(* IEC 61131-3 sources: daoli-st-library/DL_Motion (part 17) *)

(* ---- FB_DL_ServoVelLoopBand.st ---- *)
(* ===========================================================================
   组件名   : FB_DL_ServoVelLoopBand
   分类     : DL_Motion / 速度环带宽估算
   一句话   : 由速度指令阶跃响应的 10%→90% 上升时间估算闭环带宽并判定是否达标
   复杂度   : 2        版本 : v1.0.0        日期 : 2026-11-24
   开源溯源 : 无（clean-room 自研，未借鉴任何开源实现）
   输入契约 : xEnable 功能使能；xArm 测量许可（FALSE 复位）；fVelRef 速度指令 [rpm]
              fVelFbk 速度反馈 [rpm]；fDtSec 采样周期 [s]；fStepThr 阶跃识别阈值 [rpm]
              fRiseLowFrac/fRiseHighFrac 上升时间取点分数；fTimeoutSec 测量超时 [s]
              fBandFactor 上升时间-带宽系数（一阶近似 0.35）；fBandTargetHz 达标带宽 [Hz]
   输出契约 : fRiseTimeSec 上升时间 [s]；fBandwidthHz 估算带宽 [Hz]；xDone 测量完成
              xBandOk 带宽达标（容差比较）；xValid 输入有效
              iErrorCode 0=正常 1=输入非有限 2=测量超时 3=上升时间过小 9=非法状态
   修改记录 : v1.0.0 2026-11-24 初版
   =========================================================================== *)

TYPE E_DL_RiseMeasState :
(
    eIdle := 0,       // 空闲待命 | idle
    eWaitStep := 1,   // 等待阶跃发生 | wait for step
    eRising := 2,     // 上升沿测量中 | rising measurement
    eDone := 3,       // 测量完成 | measurement done
    eFail := 4        // 测量失败 | measurement failed
);
END_TYPE

FUNCTION_BLOCK FB_DL_ServoVelLoopBand
VAR_INPUT
    xEnable : BOOL;                       // 功能使能 | function enable
    xArm : BOOL;                          // 测量许可 FALSE=复位 | measurement arm
    fVelRef : REAL;                       // 速度指令 [rpm] | velocity reference [rpm]
    fVelFbk : REAL;                       // 速度反馈 [rpm] | velocity feedback [rpm]
    fDtSec : REAL := 0.004;               // 采样周期 [s] | sample period [s]
    fStepThr : REAL := 50.0;              // 阶跃识别阈值 [rpm] | step detect threshold [rpm]
    fRiseLowFrac : REAL := 0.1;           // 上升时间起点分数 | rise time low fraction
    fRiseHighFrac : REAL := 0.9;          // 上升时间终点分数 | rise time high fraction
    fTimeoutSec : REAL := 5.0;            // 测量超时 [s] | measurement timeout [s]
    fBandFactor : REAL := 0.35;           // 上升时间-带宽系数 | rise time band factor
    fBandTargetHz : REAL := 100.0;        // 达标带宽 [Hz] | target bandwidth [Hz]
END_VAR
VAR_OUTPUT
    fRiseTimeSec : REAL;                  // 上升时间 [s] | rise time [s]
    fBandwidthHz : REAL;                  // 估算带宽 [Hz] | estimated bandwidth [Hz]
    xDone : BOOL;                         // 测量完成 | measurement done
    xBandOk : BOOL;                       // 带宽达标 | bandwidth acceptable
    xValid : BOOL;                        // 输入有效标志 | inputs valid flag
    iErrorCode : INT;                     // 故障码 0=无故障 | error code
    eStateOut : E_DL_RiseMeasState;       // 当前状态观测 | current state observation
END_VAR
VAR
    _eState : E_DL_RiseMeasState := eIdle;  // 内部状态机状态 | internal state
    _fRefPrev : REAL;                     // 上一拍速度指令 [rpm] | previous reference [rpm]
    _fStart : REAL;                       // 阶跃起点值 [rpm] | step start value [rpm]
    _fAmp : REAL;                         // 阶跃幅值 [rpm] | step amplitude [rpm]
    _fElapsed : REAL;                     // 阶跃后累计时间 [s] | elapsed since step [s]
    _fProg : REAL;                        // 归一化响应进度 | normalized response progress
    _fT10 : REAL;                         // 10% 时刻 [s] | time at low fraction [s]
    _fT90 : REAL;                         // 90% 时刻 [s] | time at high fraction [s]
    _fDt : REAL;                          // 钳位后采样周期 [s] | clamped dt [s]
    _xGot10 : BOOL;                       // 已捕获低分数时刻 | low fraction captured
    _xGot90 : BOOL;                       // 已捕获高分数时刻 | high fraction captured
    _xBad : BOOL;                         // 输入非有限标志 | not-finite flag
    _xBadPar : BOOL;                      // 参数非法标志 | invalid parameter flag
END_VAR

// ---- 非有限检测 ----
_xBad := (fVelRef <> fVelRef) OR ((fVelRef - fVelRef) <> (fVelRef - fVelRef))
      OR (fVelFbk <> fVelFbk) OR ((fVelFbk - fVelFbk) <> (fVelFbk - fVelFbk))
      OR (fDtSec <> fDtSec) OR ((fDtSec - fDtSec) <> (fDtSec - fDtSec))
      OR (fBandFactor <> fBandFactor) OR ((fBandFactor - fBandFactor) <> (fBandFactor - fBandFactor));

// ---- 参数合法性：所有做分母/做取点的量必须为正且分数有序 ----
_xBadPar := (fDtSec <= 0.0) OR (fStepThr <= 0.0) OR (fTimeoutSec <= 0.0)
         OR (fBandFactor <= 0.0) OR (fBandTargetHz <= 0.0)
         OR (fRiseLowFrac <= 0.0) OR (fRiseHighFrac <= fRiseLowFrac);

xValid := NOT (_xBad OR _xBadPar);
iErrorCode := 0;
IF _xBad THEN
    iErrorCode := 1;
ELSIF _xBadPar THEN
    iErrorCode := 2;
END_IF

// ---- 周期钳位 ----
_fDt := fDtSec;
IF _fDt < 0.000001 THEN
    _fDt := 0.000001;
ELSIF _fDt > 0.2 THEN
    _fDt := 0.2;
END_IF

CASE _eState OF
    eIdle:
        xDone := FALSE;
        IF NOT xEnable THEN
            iErrorCode := 0;
        ELSIF xArm AND xValid THEN
            fRiseTimeSec := 0.0;
            fBandwidthHz := 0.0;
            xBandOk := FALSE;
            _fElapsed := 0.0;
            _eState := eWaitStep;
        END_IF

    eWaitStep:
        IF NOT xArm OR NOT xEnable THEN
            _eState := eIdle;
        ELSIF ABS(fVelRef - _fRefPrev) > fStepThr THEN
            _fStart := _fRefPrev;                    // 阶跃起点
            _fAmp := fVelRef - _fRefPrev;            // 阶跃幅值
            IF ABS(_fAmp) > 0.000000001 THEN          // 防零除：幅值必须显著
                _fElapsed := 0.0;
                _fT10 := 0.0;
                _fT90 := 0.0;
                _xGot10 := FALSE;
                _xGot90 := FALSE;
                _eState := eRising;
            ELSE
                iErrorCode := 3;                     // 幅值过小视为无效阶跃
                _eState := eFail;
            END_IF
        END_IF

    eRising:
        IF NOT xArm OR NOT xEnable THEN
            _eState := eIdle;
        ELSE
            _fElapsed := _fElapsed + _fDt;
            _fProg := 0.0;
            IF ABS(_fAmp) > 0.000000001 THEN
                _fProg := (fVelFbk - _fStart) / _fAmp;   // 归一化进度，分母已守卫
            END_IF
            IF NOT _xGot10 AND (_fProg >= fRiseLowFrac) THEN
                _fT10 := _fElapsed;
                _xGot10 := TRUE;
            END_IF
            IF _xGot10 AND NOT _xGot90 AND (_fProg >= fRiseHighFrac) THEN
                _fT90 := _fElapsed;
                _xGot90 := TRUE;
            END_IF
            IF _xGot90 THEN
                fRiseTimeSec := _fT90 - _fT10;
                IF fRiseTimeSec > 0.000001 THEN
                    fBandwidthHz := fBandFactor / fRiseTimeSec;   // 分母已守卫
                    xDone := TRUE;
                    _eState := eDone;
                ELSE
                    iErrorCode := 3;                 // 上升时间过小，估算不可信
                    _eState := eFail;
                END_IF
            ELSIF _fElapsed > fTimeoutSec THEN
                iErrorCode := 2;                     // 响应未达 90%，测量超时
                _eState := eFail;
            END_IF
        END_IF

    eDone:
        IF NOT xArm OR NOT xEnable THEN
            xDone := FALSE;
            _eState := eIdle;                        // 结果保持至下一次重新测量
        END_IF

    eFail:
        xDone := FALSE;
        IF NOT xArm OR NOT xEnable THEN
            iErrorCode := 0;
            _eState := eIdle;
        END_IF

ELSE
    iErrorCode := 9;                                 // 非法状态兜底
    xDone := FALSE;
    _eState := eIdle;
END_CASE;

// ---- 达标判定：仅在测量完成后用容差比较带宽 ----
IF _eState = eDone THEN
    xBandOk := (fBandwidthHz + 0.000001) >= fBandTargetHz;
END_IF

_fRefPrev := fVelRef;                                // 指令历史留到拍末更新
eStateOut := _eState;
END_FUNCTION_BLOCK

(* ---- FB_DL_SingleAxis.st ---- *)
(*==============================================================================
 * 组件名称 (Component)  : FB_DL_SingleAxis
 * 所属子库 (Sublibrary) : DL_Motion
 * 当前版本 (Version)    : 1.0.0
 * 组件分类 (Category)   : 功能块（FUNCTION_BLOCK）· 单轴运动控制 · PLCopen 状态机
 * 兼容性   (Platform)   : CODESYS 3.5 / TwinCAT 3 / 汇川 InoProShop / Schneider
 *                         Machine Expert；仅依赖 Standard.library，零厂商方言
 * 功能描述 (Function)   : 实现 I_DL_MotionAxis 的单轴运动控制功能块，内含
 *                         PLCopen 轴状态机语义（eDisabled + 六态）的
 *                         clean-room 实现。bUseVirtualKinematics=TRUE 时
 *                         位置由内部梯形段积分器生成（仿真）；FALSE 时位置
 *                         直接取上层每拍注入值（真实驱动），同一状态机适配
 *                         两种模式。
 * 设计要点 (Key notes)  : ① 指令仲裁 Absolute>Relative>Velocity，落选者丢弃
 *                           置信息级 0101；eStopping/eErrorStop 拒绝一切运动
 *                           指令（MC_Stop 语义）；
 *                         ② 软限位越限预判拦截（0202）；驱动故障 → eErrorStop
 *                           锁存（R15，仅 Reset 清）；非法状态 CASE+ELSE 兜底
 *                           （0201）；
 *                         ③ bError 派生式仅反映 eErrorStop，信息级码只进
 *                           uErrorId（R21）；
 *                         ④ 首扫/跟踪判据唯一合法范式 IF bTrack OR (NOT bInit)
 *                           （R5 公约 0.1）：中途跟踪脉冲 → 位置重同步并受控
 *                           停车（验收向量 V3）。
 * 输出实现 (Out mapping): 规格引脚表 OUT 列以接口 PROPERTY GET 形式实现并
 *                         与引脚表一一对应（接口契约映射），避免接口属性与
 *                         同名输出变量在编译器内重名冲突。
 * 开源溯源 (Origin)     : plcopen / s7-motion。仅提取 PLCopen 轴状态机公开
 *                         状态语义与 S7-1500 Motion Control 手册公开参数域；
 *                         状态机与梯形积分 100% 自有 clean-room，未调用任何
 *                         厂商轴控功能块，未参考任何厂商源码行。
 * 验收向量 (Acceptance) :
 *   V1 正常链：Enable→eStandstill→MoveAbsolute(120)→eDiscreteMotion→到位回
 *      eStandstill，fPosition 终值 120±0.01；
 *   V2 非法态兜底：内部状态破坏 → CASE+ELSE 兜底 → eErrorStop，码 0004_0201；
 *   V3 中途插入跟踪脉冲：bTrack=TRUE 一拍 → 位置重同步 fActPosition，运动转
 *      eStopping（0.1 公约必测向量）；V4~V6：仲裁丢弃 0101 / 目标超限拒绝
 *      0202 / 驱动故障锁存 0203 仅 Reset 可清。
 * 故障码表 (Error codes):
 *   16#0004_0101/0103/0104/0105【信息级】指令仲裁丢弃 / 参数对调兜底修复 /
 *   采样周期钳位 / 软限位预判降速停车；16#0004_0201/0202/0203【故障级】
 *   非法状态兜底 / 软限位越界（目标拒绝为瞬态码，实际越限为锁存）/
 *   驱动故障反馈锁存。
 * 修订历史 (Revision)   :
 *   2026-11-15  v1.0.0  首版入库（Round 05 · DL_Motion 开库）
 *============================================================================*)
(* 调用示例：fbAxis.fSoftLimitPos := 800.0（组态期赋值）；周期调用
 * fbAxis(bUseVirtualKinematics := TRUE, bDriveReady := TRUE)；真实驱动模式
 * 下层每拍写 fActPosition；HMI 取状态经属性 eState / fPosition / uErrorId。 *)
FUNCTION_BLOCK FB_DL_SingleAxis IMPLEMENTS I_DL_MotionAxis
VAR_INPUT
    fSoftLimitPos         : REAL := 1000000.0;  // 软限位上限（Soft limit positive）[mm]，默认 +1E6
    fSoftLimitNeg         : REAL := -1000000.0; // 软限位下限（Soft limit negative）[mm]，默认 -1E6
    fVelMax               : REAL := 1000.0;     // 速度物理上限（Max velocity）[mm/s]
    fAccMax               : REAL := 10000.0;    // 加速度物理上限（Max acceleration）[mm/s²]
    fDecMax               : REAL := 10000.0;    // 减速度物理上限（Max deceleration）[mm/s²]
    fPosTolerance         : REAL := 0.01;       // 到位容差（Position tolerance）[mm]
    tSampleTime           : TIME := T#100MS;    // 虚拟积分采样周期（Sample time），<T#10MS 钳位（公约 0.5）
    bDriveReady           : BOOL := FALSE;      // 驱动就绪反馈（Drive ready feedback），TRUE=可上使能
    bDriveFault           : BOOL := FALSE;      // 驱动故障反馈（Drive fault feedback），TRUE=故障
    fActPosition          : REAL := 0.0;        // 实际位置注入（Actual position injection）[mm]，真实驱动由上层每拍写入
    bUseVirtualKinematics : BOOL := TRUE;       // 虚拟运动学开关（Virtual kinematics），TRUE=无硬件仿真模式
    bTrack                : BOOL := FALSE;      // 跟踪脉冲（Tracking pulse），电平生效重同步位置（R5 公约 0.1）
END_VAR
VAR
    bInit                 : BOOL := FALSE;      // 首扫标志（First-scan flag，R19 范式配套）
    bReqEnable            : BOOL := FALSE;      // 使能电平请求（Enable level request）
    bReqReset             : BOOL := FALSE;      // 复位单发请求（Reset pulse request）
    bReqStop              : BOOL := FALSE;      // 停止单发请求（Stop pulse request）
    bReqMoveAbs           : BOOL := FALSE;      // 绝对定位单发请求（MoveAbsolute pulse request）
    bReqMoveRel           : BOOL := FALSE;      // 相对定位单发请求（MoveRelative pulse request）
    bReqMoveVel           : BOOL := FALSE;      // 速度模式单发请求（MoveVelocity pulse request）
    _eState               : E_DL_AxisState := E_DL_AxisState.eDisabled; // 内部状态机步序（Internal axis state）
    _fPosition            : REAL := 0.0;        // 内部当前位置（Internal position）[mm]
    _fVelocity            : REAL := 0.0;        // 内部当前速度（Internal velocity）[mm/s]
    _bEnabled             : BOOL := FALSE;      // 内部使能标志（Internal enabled flag）
    _bHomed               : BOOL := FALSE;      // 内部回原标志（Internal homed flag），本轮占位 FALSE
    _bError               : BOOL := FALSE;      // 内部故障派生位（Internal derived error flag）
    _uErrorId             : UDINT := 0;         // 内部末次事件码（Internal last error code）
    fTgtPosition          : REAL := 0.0;        // 定位目标位置（Target position）[mm]
    fRelDist              : REAL := 0.0;        // 相对位移暂存（Relative distance buffer）[mm]
    fTgtVelocity          : REAL := 0.0;        // 目标速度幅值（Target speed magnitude）[mm/s]，恒正
    fTgtVelSigned         : REAL := 0.0;        // 速度模式带符号目标（Signed velocity target）[mm/s]
    fTgtAccel             : REAL := 0.0;        // 生效加速度（Effective acceleration）[mm/s²]
    fTgtDecel             : REAL := 0.0;        // 生效减速度（Effective deceleration）[mm/s²]
    fVelCmd               : REAL := 0.0;        // 带符号速度指令（Signed velocity command）[mm/s]
    fLimPos               : REAL := 1000000.0;  // 生效软限位上限（Effective soft limit high）[mm]
    fLimNeg               : REAL := -1000000.0; // 生效软限位下限（Effective soft limit low）[mm]
    fVelLim               : REAL := 1000.0;     // 生效速度上限（Effective velocity limit）[mm/s]
    fAccLim               : REAL := 10000.0;    // 生效加速度上限（Effective acceleration limit）[mm/s²]
    fDecLim               : REAL := 10000.0;    // 生效减速度上限（Effective deceleration limit）[mm/s²]
    fDt                   : REAL := 0.1;        // 生效采样周期（Effective sample time）[s]
    fDelta                : REAL := 0.0;        // 剩余位移中间量（Remaining distance）[mm]
    fDir                  : REAL := 1.0;        // 运动方向系数（Direction factor）[1]，+1/-1
    fStopDist             : REAL := 0.0;        // 当前速度制动距离（Braking distance）[mm]
    fDistToLim            : REAL := 0.0;        // 沿运动方向距限位距离（Distance to limit）[mm]
    fVelMag               : REAL := 0.0;        // 速度幅值中间量（Velocity magnitude temp）[mm/s]
    bCmdAbsArb            : BOOL := FALSE;      // 仲裁胜出：绝对定位（Arbitration winner: absolute）
    bCmdRelArb            : BOOL := FALSE;      // 仲裁胜出：相对定位（Arbitration winner: relative）
    bCmdVelArb            : BOOL := FALSE;      // 仲裁胜出：速度模式（Arbitration winner: velocity）
    rtrigReqAbs           : R_TRIG;             // 绝对定位请求沿检测（Rising edge of MoveAbsolute request）
    rtrigReqRel           : R_TRIG;             // 相对定位请求沿检测（Rising edge of MoveRelative request）
    rtrigReqVel           : R_TRIG;             // 速度模式请求沿检测（Rising edge of MoveVelocity request）
    rtrigReqStop          : R_TRIG;             // 停止请求沿检测（Rising edge of Stop request）
    rtrigReqReset         : R_TRIG;             // 复位请求沿检测（Rising edge of Reset request）
END_VAR
VAR CONSTANT
    DL_AX_INF_MAX         : REAL := 1.0E30;     // 有限值判定幅值上限（Finite-value magnitude bound）[mm]
    DL_AX_EPS             : REAL := 1.0E-6;     // 浮点判零容差（Float zero tolerance）
    DL_AX_VEL_FLOOR       : REAL := 1.0E-3;     // 速度完成判据下限（Velocity completion floor）[mm/s]
    DL_AX_PARAM_FLOOR     : REAL := 1.0E-3;     // 动态参数下限兜底（Dynamic parameter floor）[mm/s 或 mm/s²]
    DL_AX_DT_MIN          : REAL := 0.010;      // 采样周期钳位下限（Sample time clamp low）[s]
    DL_AX_DT_MAX          : REAL := 1.0;        // 采样周期钳位上限（Sample time clamp high）[s]
END_VAR

METHOD Enable : BOOL
VAR_INPUT
    bOn : BOOL;                                  // 使能电平（Enable on/off），TRUE=上使能请求
END_VAR
IF bOn AND ((_eState = E_DL_AxisState.eErrorStop) OR bDriveFault OR (NOT bDriveReady)) THEN
    Enable := FALSE;                             // 故障/未就绪拒绝上使能（MC_Power 语义）
ELSE
    bReqEnable := bOn;
    Enable := TRUE;
END_IF
    END_METHOD

METHOD Reset : BOOL
VAR_INPUT
END_VAR
Reset := FALSE;
IF _eState = E_DL_AxisState.eErrorStop THEN
    bReqReset := TRUE;                           // 复位请求单发化，主体 eErrorStop 分支消费
    Reset := TRUE;
END_IF
    END_METHOD

METHOD Stop
VAR_INPUT
END_VAR
IF _bEnabled AND (_eState <> E_DL_AxisState.eErrorStop) THEN
    bReqStop := TRUE;                            // MC_Stop 语义：受控停车并拒绝新任务
END_IF
    END_METHOD

METHOD MoveAbsolute : BOOL
VAR_INPUT
    fPos : REAL;                                 // 目标绝对位置（Target absolute position）[mm]
    fVel : REAL;                                 // 运行速度（Run velocity）[mm/s]，正值
    fAcc : REAL;                                 // 加/减速度（Acceleration and deceleration）[mm/s²]，正值
END_VAR
MoveAbsolute := FALSE;
IF _eState <> E_DL_AxisState.eStandstill THEN RETURN; END_IF  // 非待机态拒绝
IF (fPos <> fPos) OR (fVel <> fVel) OR (fAcc <> fAcc) OR (ABS(fPos) > DL_AX_INF_MAX)
   OR (fVel <= DL_AX_PARAM_FLOOR) OR (fAcc <= DL_AX_PARAM_FLOOR) THEN RETURN; END_IF  // 参数非法/非有限值拒绝（0.8 公约）
IF (fPos > fLimPos) OR (fPos < fLimNeg) THEN
    _uErrorId := 16#0004_0202;                   // 软限位预判拦截：目标位超限直接拒绝
    RETURN;
END_IF
fTgtPosition := fPos;  fTgtVelocity := MIN(fVel, fVelLim);           // 目标位置 [mm] / 速度钳位 [mm/s]
fTgtAccel := MIN(fAcc, fAccLim);  fTgtDecel := MIN(fAcc, fDecLim);   // 加/减速度钳位 [mm/s²]
bReqMoveAbs := TRUE;
MoveAbsolute := TRUE;
    END_METHOD

METHOD MoveRelative : BOOL
VAR_INPUT
    fDist : REAL;                                // 相对位移（Relative distance）[mm]，带符号
    fVel  : REAL;                                // 运行速度（Run velocity）[mm/s]，正值
    fAcc  : REAL;                                // 加/减速度（Acceleration and deceleration）[mm/s²]，正值
END_VAR
MoveRelative := FALSE;
IF _eState <> E_DL_AxisState.eStandstill THEN RETURN; END_IF
IF (fDist <> fDist) OR (fVel <> fVel) OR (fAcc <> fAcc) OR (ABS(fDist) > DL_AX_INF_MAX)
   OR (fVel <= DL_AX_PARAM_FLOOR) OR (fAcc <= DL_AX_PARAM_FLOOR) THEN RETURN; END_IF  // 参数非法/非有限值拒绝（0.8 公约）
IF (_fPosition + fDist > fLimPos) OR (_fPosition + fDist < fLimNeg) THEN
    _uErrorId := 16#0004_0202;                   // 相对目标落点越限拒绝（预判）
    RETURN;
END_IF
fRelDist := fDist;  fTgtVelocity := MIN(fVel, fVelLim);              // 相对位移暂存 [mm] / 速度钳位
fTgtAccel := MIN(fAcc, fAccLim);  fTgtDecel := MIN(fAcc, fDecLim);
bReqMoveRel := TRUE;
MoveRelative := TRUE;
    END_METHOD

METHOD MoveVelocity : BOOL
VAR_INPUT
    fVel : REAL;                                 // 目标速度（Target velocity）[mm/s]，带符号
    fAcc : REAL;                                 // 加/减速度（Acceleration and deceleration）[mm/s²]，正值
END_VAR
MoveVelocity := FALSE;
IF (_eState <> E_DL_AxisState.eStandstill) AND (_eState <> E_DL_AxisState.eContinuousMotion) THEN
    RETURN;                                      // 待机/连续运动两态可进（连续运动中允许改速）
END_IF
IF (fVel <> fVel) OR (fAcc <> fAcc) OR (fAcc <= DL_AX_PARAM_FLOOR) THEN RETURN; END_IF
fTgtVelSigned := MAX(MIN(fVel, fVelLim), -fVelLim);  // 带符号速度钳位 [mm/s]
fTgtAccel := MIN(fAcc, fAccLim);  fTgtDecel := MIN(fAcc, fDecLim);
bReqMoveVel := TRUE;
MoveVelocity := TRUE;
(* 属性实现（PROPERTY GET）：与规格引脚表 OUT 列一一对应（接口契约映射）。 *)
    END_METHOD

// 段 1｜沿检测与单发化消费：R_TRIG 无条件周期刷新（R7 红线），标志本拍即清
rtrigReqAbs(CLK := bReqMoveAbs);  rtrigReqRel(CLK := bReqMoveRel);
rtrigReqVel(CLK := bReqMoveVel);  rtrigReqStop(CLK := bReqStop);
rtrigReqReset(CLK := bReqReset);
IF bReqMoveAbs THEN bReqMoveAbs := FALSE; END_IF   // 防标志滞留丢边沿
IF bReqMoveRel THEN bReqMoveRel := FALSE; END_IF
IF bReqMoveVel THEN bReqMoveVel := FALSE; END_IF
IF bReqStop THEN bReqStop := FALSE; END_IF
IF bReqReset THEN bReqReset := FALSE; END_IF

// 段 2｜R19 首扫/跟踪同步：判据唯一合法范式 IF bTrack OR (NOT bInit)
IF bTrack OR (NOT bInit) THEN
    IF (fActPosition = fActPosition) AND (ABS(fActPosition) <= DL_AX_INF_MAX) THEN _fPosition := fActPosition; END_IF // 位置重同步 [mm]
    fVelCmd := 0.0;                              // 首扫/跟踪清除速度指令 [mm/s]
    IF bInit AND ((_eState = E_DL_AxisState.eDiscreteMotion) OR (_eState = E_DL_AxisState.eContinuousMotion)) THEN
        _eState := E_DL_AxisState.eStopping;     // 中途插入跟踪脉冲 → 受控停车（验收向量 V3）
    END_IF
    bInit := TRUE;
END_IF

// 段 3｜参数防御与对调自修复（公约 0.6/0.8）：信息级码，不置 _bError（R21）
IF fSoftLimitPos < fSoftLimitNeg THEN
    fLimPos := fSoftLimitNeg;  fLimNeg := fSoftLimitPos;  _uErrorId := 16#0004_0103; // 对调修复
ELSE
    fLimPos := fSoftLimitPos;  fLimNeg := fSoftLimitNeg;
END_IF
IF (fVelMax > DL_AX_PARAM_FLOOR) AND (fVelMax < DL_AX_INF_MAX) THEN fVelLim := fVelMax;
ELSE fVelLim := 1000.0;  _uErrorId := 16#0004_0103; END_IF   // 非法速度上限兜底 [mm/s]
IF (fAccMax > DL_AX_PARAM_FLOOR) AND (fAccMax < DL_AX_INF_MAX) THEN fAccLim := fAccMax;
ELSE fAccLim := 10000.0;  _uErrorId := 16#0004_0103; END_IF  // 非法加速度上限兜底 [mm/s²]
IF (fDecMax > DL_AX_PARAM_FLOOR) AND (fDecMax < DL_AX_INF_MAX) THEN fDecLim := fDecMax;
ELSE fDecLim := 10000.0;  _uErrorId := 16#0004_0103; END_IF  // 非法减速度上限兜底 [mm/s²]
IF tSampleTime < T#10MS THEN fDt := DL_AX_DT_MIN;  _uErrorId := 16#0004_0104;   // 周期下限钳位 [s]
ELSIF tSampleTime > T#1S THEN fDt := DL_AX_DT_MAX;  _uErrorId := 16#0004_0104;  // 周期上限钳位 [s]
ELSE fDt := TIME_TO_REAL(tSampleTime) / 1000.0; END_IF                           // 合法周期换算 [s]

// 段 4｜驱动故障最高优先级锁存（R15：仅 Reset 可清）
IF bDriveFault THEN _eState := E_DL_AxisState.eErrorStop;  _uErrorId := 16#0004_0203; END_IF

// 段 5｜停止请求前置处理（MC_Stop 语义：使能运动/静止态均可进入停止）
IF rtrigReqStop.Q AND _bEnabled AND (_eState <> E_DL_AxisState.eStopping)
   AND (_eState <> E_DL_AxisState.eErrorStop) THEN
    _eState := E_DL_AxisState.eStopping;
END_IF

// 段 6｜同拍多指令仲裁：Absolute > Relative > Velocity，落选者丢弃
bCmdAbsArb := rtrigReqAbs.Q AND (_eState = E_DL_AxisState.eStandstill);
bCmdRelArb := (NOT bCmdAbsArb) AND rtrigReqRel.Q AND (_eState = E_DL_AxisState.eStandstill);
bCmdVelArb := (NOT bCmdAbsArb) AND (NOT bCmdRelArb) AND rtrigReqVel.Q
             AND ((_eState = E_DL_AxisState.eStandstill) OR (_eState = E_DL_AxisState.eContinuousMotion));
IF (rtrigReqAbs.Q AND (rtrigReqRel.Q OR rtrigReqVel.Q)) OR (rtrigReqRel.Q AND rtrigReqVel.Q) THEN
    _uErrorId := 16#0004_0101;                   // 信息级：指令丢弃提示（R21：不置故障）
END_IF

// 段 7｜PLCopen 轴状态机（ENUM + CASE + ELSE 兜底）
CASE _eState OF
    E_DL_AxisState.eDisabled:                    // 禁用态：等待上使能
        _bEnabled := FALSE;
        fVelCmd := 0.0;
        IF bReqEnable AND bDriveReady AND (NOT bDriveFault) THEN _bEnabled := TRUE;  _eState := E_DL_AxisState.eStandstill; END_IF
    E_DL_AxisState.eStandstill:                  // 待机态：接收运动指令
        IF NOT bReqEnable THEN
            _eState := E_DL_AxisState.eDisabled; // 下使能
        ELSIF bCmdAbsArb THEN _eState := E_DL_AxisState.eDiscreteMotion;
        ELSIF bCmdRelArb THEN
            fTgtPosition := _fPosition + fRelDist;         // 相对目标落位时现算 [mm]
            IF (fTgtPosition > fLimPos) OR (fTgtPosition < fLimNeg) THEN _uErrorId := 16#0004_0202; // 目标越限拒绝（瞬态码）
            ELSE _eState := E_DL_AxisState.eDiscreteMotion; END_IF
        ELSIF bCmdVelArb THEN _eState := E_DL_AxisState.eContinuousMotion;
        END_IF
    E_DL_AxisState.eDiscreteMotion:              // 离散运动：梯形速度规划（简化 S 曲线思想）
        fDelta := fTgtPosition - _fPosition;
        IF (ABS(fDelta) <= fPosTolerance) AND (ABS(fVelCmd) <= DL_AX_VEL_FLOOR) THEN
            fVelCmd := 0.0;                      // 到位：容差 + 速度收敛双判据
            _eState := E_DL_AxisState.eStandstill;
        ELSE
            fDir := 1.0;
            IF fDelta < 0.0 THEN fDir := -1.0; END_IF
            fStopDist := (fVelCmd * fVelCmd) / (2.0 * MAX(fTgtDecel, DL_AX_PARAM_FLOOR)); // 制动距离 [mm]，防除零
            IF fStopDist >= ABS(fDelta) THEN fVelMag := MAX(ABS(fVelCmd) - fTgtDecel * fDt, 0.0);  // 减速段 [mm/s]
            ELSE fVelMag := MIN(ABS(fVelCmd) + fTgtAccel * fDt, fTgtVelocity); END_IF              // 加速/恒速段 [mm/s]
            fVelCmd := fDir * fVelMag;
        END_IF
    E_DL_AxisState.eContinuousMotion:            // 连续运动：速度斜坡 + 软限位预判
        IF (_fPosition > fLimPos) OR (_fPosition < fLimNeg) THEN _uErrorId := 16#0004_0202;  // 实际位置越限：故障级
        _eState := E_DL_AxisState.eErrorStop;
        ELSE
            IF fTgtVelSigned > 0.0 THEN fDistToLim := fLimPos - _fPosition;    // 正向距限位 [mm]
            ELSIF fTgtVelSigned < 0.0 THEN fDistToLim := _fPosition - fLimNeg; // 负向距限位 [mm]
            ELSE fDistToLim := fPosTolerance; END_IF
            fStopDist := (fVelCmd * fVelCmd) / (2.0 * MAX(fTgtDecel, DL_AX_PARAM_FLOOR)); // 防除零
            IF fDistToLim <= fStopDist THEN
                fTgtVelSigned := 0.0;            // 预判进入警戒区 → 强制减速（信息级 0004_0105）
                _uErrorId := 16#0004_0105;
            END_IF
            IF fVelCmd < fTgtVelSigned THEN fVelCmd := MIN(fVelCmd + fTgtAccel * fDt, fTgtVelSigned);      // 速度斜坡收敛
            ELSIF fVelCmd > fTgtVelSigned THEN fVelCmd := MAX(fVelCmd - fTgtDecel * fDt, fTgtVelSigned); END_IF
            IF (ABS(fTgtVelSigned) <= DL_AX_EPS) AND (ABS(fVelCmd) <= DL_AX_VEL_FLOOR) THEN
                fVelCmd := 0.0;                  // 限位停车完成
                _eState := E_DL_AxisState.eStandstill;
            END_IF
        END_IF
    E_DL_AxisState.eStopping:                    // 受控停止：按生效减速度斜坡归零
        fVelMag := MAX(ABS(fVelCmd) - MAX(fTgtDecel, DL_AX_PARAM_FLOOR) * fDt, 0.0);
        IF fVelCmd < 0.0 THEN fVelCmd := -fVelMag; ELSE fVelCmd := fVelMag; END_IF
        IF fVelMag <= DL_AX_VEL_FLOOR THEN fVelCmd := 0.0;  _eState := E_DL_AxisState.eStandstill; END_IF  // 停稳
    E_DL_AxisState.eHoming:                      // 预留态：回原序列由后续轮次 FB_DL_AxisHomingSeq 承载
        IF NOT bReqEnable THEN _eState := E_DL_AxisState.eDisabled; END_IF  // 防御驻留：仅下使能退出
    E_DL_AxisState.eErrorStop:                   // 故障停机：报警锁存，仅 Reset 可退回
        fVelCmd := 0.0;
        _bEnabled := FALSE;
        IF rtrigReqReset.Q AND (NOT bDriveFault) THEN
            _uErrorId := 0;                      // 复位清码
            IF bReqEnable AND bDriveReady THEN _eState := E_DL_AxisState.eStandstill;   // 使能保持回待机
            ELSE _eState := E_DL_AxisState.eDisabled; END_IF                            // 否则回禁用
        END_IF

    ELSE
        // 非法状态兜底（故障级）
        _uErrorId := 16#0004_0201;  _eState := E_DL_AxisState.eErrorStop;
END_CASE

// 段 8｜位置/速度出口：虚拟积分与真实注入共用同一状态机
IF bUseVirtualKinematics THEN
    _fPosition := _fPosition + fVelCmd * fDt;    // 虚拟运动学：位置积分 [mm]
ELSIF (fActPosition = fActPosition) AND (ABS(fActPosition) <= DL_AX_INF_MAX) THEN
    _fPosition := fActPosition;                  // 真实驱动：上层每拍注入 [mm]
END_IF                                           // 非有限值注入 → 保持上一拍位置（0.8 公约）
_fVelocity := fVelCmd;                           // 速度出口 = 带符号速度指令 [mm/s]
_bError := (_eState = E_DL_AxisState.eErrorStop); // bError 派生式（R21：信息级码不进 bError）

(*-----------------------------------------------------------------------------
 * 方法实现（METHOD）：全部非阻塞，仅置内部请求标志，跨周期动作由主体状态机
 * 执行（OOP 方法设计准则）；接口方法共 6 个达红线临界，不得再增。
 *-----------------------------------------------------------------------------*)

PROPERTY eState : E_DL_AxisState
eState := _eState;
END_PROPERTY
PROPERTY fPosition : REAL
fPosition := _fPosition;
END_PROPERTY
PROPERTY fVelocity : REAL
fVelocity := _fVelocity;
END_PROPERTY
PROPERTY bEnabled : BOOL
bEnabled := _bEnabled;
END_PROPERTY
PROPERTY bHomed : BOOL
bHomed := _bHomed;
END_PROPERTY
PROPERTY bError : BOOL
bError := _bError;
END_PROPERTY
PROPERTY uErrorId : UDINT
uErrorId := _uErrorId;
END_PROPERTY
END_FUNCTION_BLOCK

(* ---- FB_DL_SocketPressTrend.st ---- *)
// =====================================================================
// FB_DL_SocketPressTrend.st
// 压装压力-位移曲线特征提取与包络判定（峰值/位移窗/刚度 → OK·NG）
// Press force-position curve feature extraction and envelope FB
// 码位: 16#0004_034F ~ 16#0004_0353 (本件独占 5 槽)
// 修改记录: R29 初版 (按 DISPATCH_R29 序 15)
// =====================================================================
FUNCTION_BLOCK FB_DL_SocketPressTrend
VAR_INPUT
    bEnable       : BOOL  := FALSE;    // 使能 / Enable
    bPressStart   : BOOL  := FALSE;    // 上升沿开始采集一次 / Press start on edge
    bPressDone    : BOOL  := FALSE;    // 压装到行程结束 / Press done
    fForce_N      : REAL  := 0.0;      // 实时压力 0~50000 N / Force [N]
    fPos_mm       : REAL  := 0.0;      // 实时位移 0~200 mm / Position [mm]
    fForceMin_N   : REAL  := 500.0;    // 压力下限 >0 N / Min force [N]
    fForceMax_N   : REAL  := 5000.0;   // 压力上限 >下限 N / Max force [N]
    fPosWinLo_mm  : REAL  := 2.0;      // 峰值位移窗下限 ≥0 mm / Position window low [mm]
    fPosWinHi_mm  : REAL  := 8.0;      // 峰值位移窗上限 >下限 mm / Position window high [mm]
    fStiffMin_Nmm : REAL  := 200.0;    // 刚度下限 ≥0 N/mm / Min stiffness [N/mm]
    fReboundPct   : REAL  := 20.0;     // 峰值后取段百分比 5~50 % / Rebound segment [%]
END_VAR
VAR_OUTPUT
    fForcePeak_N  : REAL;              // 峰值压力 N / Peak force [N]
    fPosAtPeak_mm : REAL;              // 峰值处位移 mm / Position at peak [mm]
    fStiff_Nmm    : REAL;              // 刚度估计 N/mm / Stiffness [N/mm]
    bCurveOk      : BOOL;              // 曲线判 OK / Curve OK
    uCurveCnt     : UDINT;             // 已判定曲线数 / Judged curve count
    uNgCode       : USINT;             // NG 码 0=OK 1=低压 2=高压 3=位移窗 4=刚度 / NG code
    eErr          : UDINT;             // 错误码 / Error code
END_VAR
VAR
    rtrigStart    : R_TRIG;            // 启动沿检测（无条件刷新）/ Start edge detector
    rtrigDone     : R_TRIG;            // 完成沿检测（无条件刷新）/ Done edge detector
    aForceBuf     : ARRAY[0..511] OF REAL;     // 压力采集缓冲 / Force capture buffer [N]
    aPosBuf       : ARRAY[0..511] OF REAL;     // 位移采集缓冲 / Position capture buffer [mm]
    uSampleCnt    : UDINT;             // 已采样点数 / Sample count
    uIdx          : UDINT;             // 循环下标 / Loop index
    uK            : INT;               // 采样下标 / Sample subscript
    bCollecting   : BOOL  := FALSE;    // 采集中 / Collecting flag
    bJudged       : BOOL  := FALSE;    // 本曲线已结算 / Judged flag
    bStarted      : BOOL  := FALSE;    // 曾收到启动沿 / Ever started flag
    uPeakIdx      : UDINT;             // 峰值采样序号 / Peak sample index
    fForceLimit   : REAL;              // 峰值后回弹取段力阈 / Rebound segment force threshold [N]
    fReboundHi    : REAL;              // 回弹区间位移上界 / Rebound position upper [mm]
    fPosRef       : REAL;              // 刚度段参考位移 / Stiffness reference position [mm]
    fFRef         : REAL;              // 刚度段参考力 / Stiffness reference force [N]
    fDPos         : REAL;              // 位移差 / Position delta [mm]
    fDForce       : REAL;              // 力差 / Force delta [N]
    xFirstScan    : BOOL  := TRUE;     // 首扫标记 / First-scan flag
END_VAR

// ---------------------------------------------------------------------
// 代码位表（本件独占，勿复用）:
//   16#0004_034F 信息 曲线判定 OK
//   16#0004_0350 故障 压力/位移非有限
//   16#0004_0351 故障 fForceMax_N ≤ fForceMin_N / fPosWinHi_mm ≤ fPosWinLo_mm / fStiffMin_Nmm < 0（组态错）
//   16#0004_0352 信息 曲线 NG（bCurveOk=FALSE 且 uNgCode>0）——NG 是产品判据不是设备故障
//   16#0004_0353 信息 bPressDone 在从未收到 bPressStart 时置位（时序错）→ 丢弃本次、不出结论
// ---------------------------------------------------------------------

// ---- 沿检测（每拍无条件刷新，R7 纪律）/ Edge detection, unconditional ----
rtrigStart(CLK := bPressStart); // 启动沿 / Start edge
rtrigDone(CLK := bPressDone);   // 完成沿 / Done edge

// ---- 非有限闸 / Finite gate ----
IF (fForce_N <> fForce_N) OR (ABS(fForce_N) >= 1.0E12)
   OR (fPos_mm <> fPos_mm) OR (ABS(fPos_mm) >= 1.0E12) THEN
    eErr := 16#0004_0350;       // 故障码 / Fault code
    RETURN;                     // 采集暂停保持 / Collection holds
END_IF

// ---- 组态错闸 / Configuration fault gate ----
IF (fForceMax_N <= fForceMin_N)
   OR (fPosWinHi_mm <= fPosWinLo_mm)
   OR (fStiffMin_Nmm < 0.0)
   OR (fForceMin_N <= 0.0) THEN
    eErr := 16#0004_0351;       // 故障码 / Fault code
    RETURN;                     // 本拍结束 / End of cycle
END_IF

// ---- 首扫初始化（R16 首扫纪律）/ First-scan initialization ----
IF xFirstScan THEN
    bCurveOk := FALSE;          // 结论复位 / Verdict reset
    uNgCode := 0;               // NG 码复位 / NG code reset
    fForcePeak_N := 0.0;        // 峰值清零 / Peak cleared
    fPosAtPeak_mm := 0.0;       // 峰位清零 / Peak position cleared
    fStiff_Nmm := 0.0;          // 刚度清零 / Stiffness cleared
    xFirstScan := FALSE;        // 清标记 / Clear flag
END_IF

// ---- 使能撤销 / Disable ----
IF NOT bEnable THEN
    bCollecting := FALSE;       // 采集退出 / Collection off
    bStarted := FALSE;          // 启动历史复位 / Started reset
    eErr := 16#0004_034F;       // 信息级：空闲 / Info: idle
    RETURN;                     // 本拍结束 / End of cycle
END_IF

// ---- 时序错：未收到启动沿就收到完成沿 → 丢弃不出结论 / Sequence error: done without start ----
IF rtrigDone.Q AND (NOT bStarted) THEN
    bCollecting := FALSE;       // 采集复位 / Collection reset
    bJudged := FALSE;           // 结算标志复位 / Judged reset
    eErr := 16#0004_0353;       // 信息级：时序错 / Info: sequence error
    RETURN;                     // uCurveCnt 不变 / Count unchanged
END_IF

// ---- 启动沿：开新曲线采集 / Start edge: begin new capture ----
IF rtrigStart.Q THEN
    bCollecting := TRUE;        // 采集开始 / Collecting
    bStarted := TRUE;           // 启动历史置位 / Started set
    bJudged := FALSE;           // 结算标志复位 / Judged reset
    uSampleCnt := 0;            // 采样计数清零 / Sample count reset
    fForcePeak_N := 0.0;        // 峰值清零 / Peak cleared
    fPosAtPeak_mm := 0.0;       // 峰位清零 / Peak position cleared
    fStiff_Nmm := 0.0;          // 刚度清零 / Stiffness cleared
    bCurveOk := FALSE;          // 结论复位 / Verdict reset
    uNgCode := 0;               // NG 码复位 / NG code reset
END_IF

// ---- 采集路径 / Collection path ----
IF bCollecting AND (NOT bJudged) THEN
    // 缓冲上限 512 点（到限停止记录并置槽 4，不覆盖前段）/ Buffer cap 512
    IF uSampleCnt < 512 THEN
        uSampleCnt := uSampleCnt + 1;   // 计数 / Count
        aForceBuf[UDINT_TO_INT(uSampleCnt - 1)] := fForce_N;    // 存力 / Store force
        aPosBuf[UDINT_TO_INT(uSampleCnt - 1)] := fPos_mm;       // 存位移 / Store position
        // 峰值跟踪 / Peak tracking
        IF fForce_N > fForcePeak_N THEN
            fForcePeak_N := fForce_N;           // 更新峰值 / Update peak
            fPosAtPeak_mm := fPos_mm;           // 峰位 / Peak position
            uPeakIdx := uSampleCnt - 1;         // 峰序号 / Peak index
        END_IF
    ELSE
        eErr := 16#0004_0352;       // 信息级：缓冲满登记 / Info: buffer full
    END_IF
END_IF

// ---- 完成沿结算（同一曲线不重复结算）/ Done edge: settle once ----
IF rtrigDone.Q AND bStarted AND (NOT bJudged) THEN
    bJudged := TRUE;            // 结算标志 / Judged set
    bCollecting := FALSE;       // 采集结束 / Collection off
    uCurveCnt := uCurveCnt + 1; // 判定计数 / Count increment

    // ---- 空压/漏装独立判：峰值 < 下限 → NG 码 1 / Under-force: NG 1 ----
    IF fForcePeak_N < fForceMin_N THEN
        bCurveOk := FALSE;      // NG / Not OK
        uNgCode := 1;           // 低压码 / Low force code
        eErr := 16#0004_0352;   // 信息级：NG / Info: NG
        RETURN;                 // 结算完成返回 / Settled
    END_IF

    // ---- 高压判 → NG 码 2 / Over force: NG 2 ----
    IF fForcePeak_N > fForceMax_N THEN
        bCurveOk := FALSE;      // NG / Not OK
        uNgCode := 2;           // 高压码 / High force code
        eErr := 16#0004_0352;   // 信息级：NG / Info: NG
        RETURN;                 // 结算完成返回 / Settled
    END_IF

    // ---- 位移窗判 → NG 码 3 / Position window: NG 3 ----
    IF (fPosAtPeak_mm < fPosWinLo_mm) OR (fPosAtPeak_mm > fPosWinHi_mm) THEN
        bCurveOk := FALSE;      // NG / Not OK
        uNgCode := 3;           // 位移窗码 / Window code
        eErr := 16#0004_0352;   // 信息级：NG / Info: NG
        RETURN;                 // 结算完成返回 / Settled
    END_IF

    // ---- 刚度估计：峰值后回弹段斜率（负斜率段不计入）/ Stiffness: rebound slope, skip negative ----
    fReboundHi := fPosWinHi_mm * 2.0;   // 搜索上界（全程扫描替代百分比近似窗）/ Search upper bound
    fPosRef := 0.0;             // 参考位移复位 / Reset ref
    fFRef := 0.0;               // 参考力复位 / Reset ref
    fStiff_Nmm := 0.0;          // 刚度复位 / Reset stiffness
    // 从峰值向后找首个有效正斜率段（回弹区间内）/ Find first valid positive slope after peak
    FOR uIdx := uPeakIdx + 1 TO uSampleCnt - 1 DO
        uK := UDINT_TO_INT(uIdx);           // 下标 / Subscript
        fDPos := aPosBuf[uK] - aPosBuf[uK - 1];     // 位移差 / Position delta
        fDForce := aForceBuf[uK] - aForceBuf[uK - 1];   // 力差 / Force delta
        IF (fDPos >= 0.01) AND (fDForce > 0.0) THEN     // 正斜率且位移够大 / Valid slope
            fStiff_Nmm := fDForce / fDPos;  // 刚度估计 / Stiffness [N/mm]
            fPosRef := aPosBuf[uK];         // 参考点 / Reference point
            fFRef := aForceBuf[uK];         // 参考力 / Reference force
        END_IF
        IF fPosRef > 0.0 THEN
            uIdx := uSampleCnt;             // 找到即提前退出扫描 / Early exit
        END_IF
    END_FOR

    // ---- 刚度判 → NG 码 4 / Stiffness: NG 4 ----
    IF fStiff_Nmm < fStiffMin_Nmm THEN
        bCurveOk := FALSE;      // NG / Not OK
        uNgCode := 4;           // 刚度码 / Stiffness code
        eErr := 16#0004_0352;   // 信息级：NG / Info: NG
        RETURN;                 // 结算完成返回 / Settled
    END_IF

    // ---- 全部通过 → OK / All passed ----
    bCurveOk := TRUE;           // OK / OK
    uNgCode := 0;               // 无 NG 码 / No NG code
    eErr := 16#0004_034F;       // 信息级：判定 OK / Info: OK
END_IF

END_FUNCTION_BLOCK

(* ---- FB_DL_SoftLimitCfgAudit.st ---- *)
(*==============================================================================
 * 组件名称 (Component)  : FB_DL_SoftLimitCfgAudit
 * 所属子库 (Sublibrary) : DL_Motion
 * 当前版本 (Version)    : 1.0.0
 * 兼容性 (Platform)     : CODESYS 3.5+ / TwinCAT 3 / 汇川 InoProShop / 施耐德 Machine Expert
 *                         仅依赖 Standard.library，零厂商私有库，零轴状态枚举（R277）
 * 功能描述 (Function)   : 软限位组态交叉审计（投运/改版期一次性或周期审计）。
 *                         对软限域 [fSoftNeg, fSoftPos]、硬限域 [fHardNeg,
 *                         fHardPos]、行程域 [fTravelNeg, fTravelPos] 做五项
 *                         交叉判定：软限域 ⊆ 硬限域（两侧）、软限域 ⊆ 行程域
 *                         （两侧）、软限间距 >= 最小有效行程；任一项不过 →
 *                         bAuditFail 锁存并逐项输出失败位（归因到项，R190 粒度）。
 *                         与 SoftLimitGuard 分工：审计组态（静态），守卫运行
 *                         （动态）。
 * 来源标签 (Origin)     : 自研线（IEC 61131-3 标准语义的道莅防御性实现，clean-room）
 * 分工声明 (Pairing)    : SoftLimitCfgAudit（组态审计，本件）↔ SoftLimitGuard
 *                         （运行守卫，既有件）：本件只判静态域包含关系，不做
 *                         运行期位置预判、不输出拦截建议（R298 属主边界）。
 * 边界语义 (Boundary)   : ① 五项判定互独立，逐项输出失败位（不合并成单一布尔
 *                         造成归因丢失，R190 口径）；
 *                         ② 域值 NaN → 对应项按失败判（审计从严：可疑组态
 *                         不得放行）；
 *                         ③ 容差比较用 DL_AUD_EPS（浮点禁等值判，R4 口径）；
 *                         ④ 组态闸：最小有效行程 < 0 → 故障锁存。
 * 输出语义 (Fallback)   : 【R191】bEnable = FALSE → 审计输出保持末值（审计
 *                         结论是台账，不随失能清零）；eFault 相 → 冻结 +
 *                         bError = TRUE。监视型无主状态机（R23 公约）。
 * 码位     (Codes)      : 按 R297 范式零 16# 码位硬编码；错误出口 BOOL+ENUM(eCause)，
 *                         码位待主控收口统一派号。
 * 红线自检 (Redline)    : 7 项红线已自检：R1 零全局 ✓｜R2 零物理地址 ✓｜R3 纯 IEC ✓
 *                         R4 NaN 从严判败/容差比较/组态闸 ✓｜R5 双语同行注释 ✓
 *                         R6 N/A（监视型无状态机，判据纯派生）✓｜R7 N/A（无实例）✓
 * 验收向量 (Acceptance) : V1 软限 [-100,100] ⊆ 硬限 [-120,120] ⊆ 行程 [-130,130]，
 *                         间距 200 >= 10 → 全过 bAuditOk=TRUE；
 *                         V2 软限正界 125 > 硬限正界 120 → bFailPosOut=TRUE；
 *                         V3 软限间距 8 < 最小行程 10 → bFailSpan=TRUE；
 *                         V4 fHardPos=NaN → bFailPosOut=TRUE（从严）。
 * 修订历史 (Revision)   : 2026-11-20  v1.0.0  R49 首版（批 4 · 序号 18）
 *==============================================================================*)
TYPE E_DL_ScaCause :
(
    eNone       := 0,                        (* 无故障成因 / No cause *)
    eCfgIllegal := 1,                        (* 组态非法：最小行程域 / Illegal config: min-span domain *)
    eAuditFail  := 2                         (* 审计不通过（失败位承载逐项归因） / Audit failed *)
);
END_TYPE

FUNCTION_BLOCK FB_DL_SoftLimitCfgAudit
VAR_INPUT
    fSoftPos    : LREAL := 100.0;            (* 软限位正界 [mm] / Soft limit positive *)
    fSoftNeg    : LREAL := (-100.0);         (* 软限位负界 [mm] / Soft limit negative *)
    fHardPos    : LREAL := 120.0;            (* 硬限位正界 [mm] / Hard limit positive *)
    fHardNeg    : LREAL := (-120.0);         (* 硬限位负界 [mm] / Hard limit negative *)
    fTravelPos  : LREAL := 130.0;            (* 机械行程正界 [mm] / Travel positive bound *)
    fTravelNeg  : LREAL := (-130.0);         (* 机械行程负界 [mm] / Travel negative bound *)
    fMinSpan    : LREAL := 10.0;             (* 软限最小有效行程要求，域 >= 0.0 [mm] / Minimum soft span requirement *)
    bRunAudit   : BOOL := FALSE;             (* 审计触发电平，TRUE 执行判定并刷新输出 [-] / Audit trigger level *)
    bReset      : BOOL := FALSE;              (* 复位命令，上升沿清审计锁存与失败位 [-] / Reset command *)
END_VAR
VAR_OUTPUT
    bAuditOk      : BOOL;                    (* 本轮审计全过电平（审计期有效）[-] / Audit-pass level *)
    bAuditFail    : BOOL;                    (* 审计不通过锁存位（复位沿清）[-] / Audit-fail latch *)
    bFailPosOutNeg: BOOL;                    (* 失败项 1：软限正界越过硬限正界 [-] / Fail item 1 *)
    bFailPosOutPos: BOOL;                    (* 失败项 2：软限负界越过硬限负界 [-] / Fail item 2 *)
    bFailTrvNeg   : BOOL;                    (* 失败项 3：软限正界越过行程正界 [-] / Fail item 3 *)
    bFailTrvPos   : BOOL;                    (* 失败项 4：软限负界越过行程负界 [-] / Fail item 4 *)
    bFailSpan     : BOOL;                    (* 失败项 5：软限间距不足最小行程 [-] / Fail item 5 *)
    nFailCnt      : INT;                     (* 本轮失败项计数 [项] / Failed item count *)
    eCause        : E_DL_ScaCause;           (* 成因出口（R190 逐项归由失败位承载） / Cause outlet *)
    bError        : BOOL;                    (* 组态故障锁存标志 [-] / Config fault flag *)
END_VAR
VAR
    rtReset   : R_TRIG;                       (* 复位沿实例，段 0 无条件调用 / Reset edge instance *)
    _bFault   : BOOL;                        (* 组态故障锁存位 / Config fault latch bit *)
    _bPosNaN  : BOOL;                        (* 任一域值非有限当拍量（从严判败用）[-] / Any bound non-finite this scan *)
    _nFail    : INT;                         (* 本轮失败项计数中间量 [项] / Fail count intermediate *)
END_VAR
VAR CONSTANT
    DL_AUD_EPS : LREAL := 1.0E-9;            (* 域比较容差（浮点禁等值判）[mm] / Domain comparison epsilon *)
END_VAR

(* —— 段 0：当拍判据派生 + 沿实例无条件刷新（R228A） —— *)
rtReset(CLK := bReset);                      (* 复位沿每拍必调 / Reset edge every scan *)
_bPosNaN := (fSoftPos <> fSoftPos) OR (fSoftNeg <> fSoftNeg) OR (fHardPos <> fHardPos)   (* 全部域值 NaN 自反判（逐引脚覆盖，R151） / NaN reflex on every bound *)
            OR (fHardNeg <> fHardNeg) OR (fTravelPos <> fTravelPos) OR (fTravelNeg <> fTravelNeg);

(* —— 段 1：复位沿处理（作用域：清故障 + 清失败锁存 + 清失败位，R283 逐项声明） —— *)
IF rtReset.Q THEN
    _bFault := FALSE;                        (* 清组态故障 / Clear fault *)
    eCause := E_DL_ScaCause.eNone;           (* 清成因 / Clear cause *)
    bAuditFail := FALSE;                     (* 清审计失败锁存 / Clear fail latch *)
    bFailPosOutNeg := FALSE;                 (* 清失败位 1 / Clear item 1 *)
    bFailPosOutPos := FALSE;                 (* 清失败位 2 / Clear item 2 *)
    bFailTrvNeg := FALSE;                    (* 清失败位 3 / Clear item 3 *)
    bFailTrvPos := FALSE;                    (* 清失败位 4 / Clear item 4 *)
    bFailSpan := FALSE;                      (* 清失败位 5 / Clear item 5 *)
    nFailCnt := 0;                           (* 清失败计数 / Clear count *)
    bAuditOk := FALSE;                       (* 清全过电平 / Clear pass level *)
END_IF

(* —— 段 2：组态闸故障锁存（最小行程负值无语义；锁存至复位沿，R189） —— *)
IF (fMinSpan < 0.0) AND NOT _bFault THEN
    _bFault := TRUE;                         (* 锁存组态故障（R45 配对） / Latch config fault *)
    eCause := E_DL_ScaCause.eCfgIllegal;     (* 成因：组态非法 / Cause: illegal config *)
END_IF

(* —— 段 3：审计判定（监视型纯派生，无 CASE 相；触发电平门控） —— *)
IF bRunAudit AND NOT _bFault THEN
    _nFail := 0;                             (* 失败计数清零重判 / Fail count recompute *)
    (* 项 1：软限正界须 < 硬限正界（从严：NaN 判败） / Item 1: soft pos must be inside hard pos *)
    IF _bPosNaN OR (fSoftPos > fHardPos - DL_AUD_EPS) THEN
        bFailPosOutNeg := TRUE;              (* 失败位 1 置位 / Item 1 fail *)
        _nFail := _nFail + 1;                (* 失败计数 / Count *)
    ELSE
        bFailPosOutNeg := FALSE;             (* 通过清位（每拍全路径赋值，R285） / Item 1 pass *)
    END_IF
    (* 项 2：软限负界须 > 硬限负界 / Item 2: soft neg inside hard neg *)
    IF _bPosNaN OR (fSoftNeg < fHardNeg + DL_AUD_EPS) THEN
        bFailPosOutPos := TRUE;              (* 失败位 2 / Item 2 fail *)
        _nFail := _nFail + 1;                (* 失败计数 / Count *)
    ELSE
        bFailPosOutPos := FALSE;             (* 通过清位 / Item 2 pass *)
    END_IF
    (* 项 3：软限正界须 <= 行程正界 / Item 3: soft pos inside travel pos *)
    IF _bPosNaN OR (fSoftPos > fTravelPos + DL_AUD_EPS) THEN
        bFailTrvNeg := TRUE;                 (* 失败位 3 / Item 3 fail *)
        _nFail := _nFail + 1;                (* 失败计数 / Count *)
    ELSE
        bFailTrvNeg := FALSE;                (* 通过清位 / Item 3 pass *)
    END_IF
    (* 项 4：软限负界须 >= 行程负界 / Item 4: soft neg inside travel neg *)
    IF _bPosNaN OR (fSoftNeg < fTravelNeg - DL_AUD_EPS) THEN
        bFailTrvPos := TRUE;                 (* 失败位 4 / Item 4 fail *)
        _nFail := _nFail + 1;                (* 失败计数 / Count *)
    ELSE
        bFailTrvPos := FALSE;                (* 通过清位 / Item 4 pass *)
    END_IF
    (* 项 5：软限间距须 >= 最小有效行程（间距 = 正界-负界，NaN 从严判败） / Item 5: span check *)
    IF _bPosNaN OR ((fSoftPos - fSoftNeg) < fMinSpan - DL_AUD_EPS) THEN
        bFailSpan := TRUE;                   (* 失败位 5 / Item 5 fail *)
        _nFail := _nFail + 1;                (* 失败计数 / Count *)
    ELSE
        bFailSpan := FALSE;                  (* 通过清位 / Item 5 pass *)
    END_IF
    nFailCnt := _nFail;                      (* 失败计数出口 / Count outlet *)
    IF _nFail > 0 THEN
        bAuditFail := TRUE;                  (* 审计失败锁存至复位沿 / Fail latch *)
        eCause := E_DL_ScaCause.eAuditFail;  (* 成因：审计不通过（逐项细节在失败位） / Cause: audit fail *)
        bAuditOk := FALSE;                   (* 全过电平收敛 / Pass level off *)
    ELSE
        bAuditOk := TRUE;                    (* 全过电平 / Pass level *)
        bAuditFail := FALSE;                 (* 通过时清失败锁存（新一轮覆盖旧结论） / Pass clears latch *)
        eCause := E_DL_ScaCause.eNone;       (* 成因清零 / Cause clear *)
    END_IF
END_IF

(* —— 段 4：出口映射（R191 名实同源） —— *)
bError := _bFault;                           (* 组态故障镜像 / Config fault mirror *)
END_FUNCTION_BLOCK

(* ---- FB_DL_SolderRibbonTension.st ---- *)
//==============================================================================
// 功能块：FB_DL_SolderRibbonTension ｜ 中文名称：焊带放卷张力与蛇形纠偏
// 所属子库：DL_Motion ｜ 版本：v1.0.0 ｜ 兼容：CODESYS V3.5+ / TwinCAT 3 / 汇川 InoProShop
// 功能描述：光伏焊带（互连条）放卷张力控制——锥度张力设定随卷径递减：
//           SP(D) = fTensionFullN x (1 - fTaperPct/100 x (D - D芯)/
//           (D满 - D芯))，卷芯处设定 = 满卷设定、满卷处设定 = 满卷设定
//           x (1 - 锥度百分比)（卷径越大张力越低，防内层压伤）；张力
//           偏差经比例修调输出（fTrimPct，给放卷驱动张力修调入口）；
//           横动机构行程窗口拦截（|位置| >= 限位即封锁横动输出）+ 接近
//           限位预警带。运行中张力 < 断带阈或 >= 超限阈（双端判据）→
//           断带/超限锁存跳闸请求。
// 开源溯源 (Origin)：道莅原创实现（参考放卷锥度张力控制工程惯例 分类与参数域）
// 单位表：张力[N] / 卷径[毫米] / 锥度[百分数] / 修调[百分数] / 修调增益
//         [百分数每牛] / 横动位置[毫米] / 时间[ms]
// 错误码表：16#0004_01E7 信息级（张力偏差进入预警带，不置 bError）/
//           16#0004_01E8 信息级（横动接近行程限位预警带，不置 bError）/
//           16#0004_0306 故障级（组态非法：卷径/张力/锥度/限位域、时间
//           窗 <= 0 或任一输入非有限，置 bError）/ 16#0004_0307 故障级
//           （断带/超限锁存：运行中张力 < 断带阈或 >= 超限阈持续去抖
//           窗，跳闸请求锁存，置 bError——该场景不可由 0306 的组态类
//           判据观测，属运行张力独立域）/ 16#0004_0308 故障级兜底（状态
//           机落 ELSE，置 bError）
// 状态机：E_DL_RibbonTenState（四态：eIdle=0 / eRun=10 / eTrip=20 /
//           eFault=99），CASE 含 ELSE 兜底，ELSE 置 0308 并撤修调输出
// 边界行为：① 组态非法 → 故障态锁存，bReset 复位；② 卷径域外钳
//           [D芯, D满] 照算（换卷瞬态照常出设定）；③ 锥度百分比域
//           [0, 100]，= 0 即恒张力；④ 横动 |位置| >= 限位 → 封锁横动
//           输出（电平），>= 90% 限位 → 信息预警；⑤ 跳闸锁存至 bReset；
//           ⑥ 安全侧 = 故障/跳闸路径修调输出撤零，禁止带故障修调。
// 修订历史：v1.0.0 2026-11-17 首版（R24 派单 · ROADMAP P1 §703）
//==============================================================================

(*------------------------------------------------------------------------------
 * 枚举: E_DL_RibbonTenState（归属本功能块，同文件发布，全库唯一定义）
 * 含义: 放卷张力相位，每个成员在 CASE 中有且仅有一个标签。
 *-----------------------------------------------------------------------------*)
TYPE E_DL_RibbonTenState :
(
    eIdle   := 0,   // 空闲：未使能 / Idle, not enabled
    eRun    := 10,  // 运行：锥度设定与修调闭环 / Run, taper setpoint and trim loop
    eTrip   := 20,  // 跳闸：断带/超限锁存 / Trip, break or over-limit latched
    eFault  := 99   // 故障：组态非法/非法状态 / Fault, config or illegal state
);
END_TYPE

FUNCTION_BLOCK FB_DL_SolderRibbonTension
VAR_INPUT
    bEnable        : BOOL;                  // 张力控制使能 [—] / Tension control enable
    bReset         : BOOL;                  // 故障复位 [—]，上升沿清锁存 / Fault reset, rising edge clears latches
    bRunning       : BOOL;                  // 放卷运行 [—]（判据与修调的使能前提） / Unwind running
    fTensionMeasN  : LREAL;                 // 张力实测 [牛] / Measured tension [N]
    fDiamNowMm     : LREAL;                 // 当前卷径 [毫米]，域外钳 [D芯, D满] 照算 / Current roll diameter [mm]
    fDiamFullMm    : LREAL := 300.0;        // 满卷直径 [毫米]，须 > 卷芯 / Full roll diameter [mm]
    fDiamCoreMm    : LREAL := 50.0;         // 卷芯直径 [毫米]，须 >= 0 且 < 满卷 / Core diameter [mm]
    fTensionFullN  : LREAL := 20.0;         // 卷芯处张力设定 [牛]，须 > 0 / Tension setpoint at the core [N]
    fTaperPct      : LREAL := 20.0;         // 锥度百分比 [百分数]，域 [0, 100]，0 = 恒张力 / Taper percent [percent], 0 = constant tension
    fTensionBreakN : LREAL := 2.0;          // 断带阈 [牛]，运行中低于此判断带 / Break threshold [N]
    fTensionOverN  : LREAL := 60.0;         // 超限阈 [牛]，运行中高于此判过张力 / Over-tension threshold [N]
    fTrimGainPctPerN: LREAL := 2.0;         // 修调增益 [百分数每牛] / Trim gain [percent/N]
    fLateralPosMm  : LREAL;                 // 横动位置 [毫米] / Lateral position [mm]
    fLateralLimitMm: LREAL := 30.0;         // 横动行程限 [毫米]，须 > 0 / Lateral travel limit [mm]
    tTripDebounce  : TIME  := T#500MS;      // 断带/超限去抖窗 [ms]，须 > 0 / Trip debounce window [ms]
END_VAR
VAR_OUTPUT
    fTensionSpN    : LREAL;                 // 锥度后张力设定 [牛]（诊断出口） / Tapered tension setpoint [N], diagnostics outlet
    fTrimPct       : LREAL;                 // 张力修调输出 [百分数]，-100..100 / Tension trim output [percent]
    bLateralBlock  : BOOL;                  // 横动封锁 [—]（行程限位电平） / Lateral block, limit level
    eState         : E_DL_RibbonTenState;   // 相位出口 [—] / Phase outlet
    eErr           : UDINT;                 // 错误码，0 = 无错，码位 16#0004_01E7 起信息级、16#0004_0306 起故障级（分带见错误码表） / Error code, 0 = no error, band info/fault per the code table
    bError         : BOOL;                  // 故障级标志，仅故障级错误置位 / Fault-class flag, set only on fault-level codes
    bValid         : BOOL;                  // 输出可用标志 / Outputs usable flag
END_VAR
VAR
    fbTrip    : TON;                        // 断带/超限去抖计时（每拍无条件刷新）[ms] / Trip debounce timer, refreshed unconditionally
    _eState   : E_DL_RibbonTenState := E_DL_RibbonTenState.eIdle; // 当前相位 / Current phase
    _bCfgBad  : BOOL;                       // 组态非法锁存 / Illegal config latch
    _bTripL   : BOOL;                       // 断带/超限锁存 / Break or over-limit latch
    _bInfoBand: BOOL;                       // 张力预警信息当拍标志 / Tension-band info flag of this scan
    _bInfoLat : BOOL;                       // 横动预警信息当拍标志 / Lateral-band info flag of this scan
    _fDiaUse  : LREAL;                      // 生效卷径（已钳位）[毫米] / Effective diameter, clamped [mm]
    _fSpanMm  : LREAL;                      // 卷径跨度 [毫米]（除零已闸） / Diameter span [mm]
    _bIllegal : BOOL;                       // 非法状态标志 / Illegal state flag
    _bInit    : BOOL := FALSE;              // 首扫标志，初值 FALSE 取非判定 / First-scan flag, tested negated
END_VAR
VAR CONSTANT
    DL_SRT_INF    : LREAL := 1.7976931348623157E308; // LREAL 幅值上限 / LREAL magnitude ceiling
    DL_SRT_EPS    : LREAL := 1.0E-6;        // 浮点判零容差 [混合] / Float zero tolerance
    DL_SRT_TRIMMAX: LREAL := 100.0;         // 修调满幅 [百分数] / Trim full scale [percent]
    DL_SRT_LATWARN: LREAL := 0.9;           // 横动预警带占比 [比值]（90% 限位） / Lateral warning ratio [ratio]
    DL_SRT_ZERO   : LREAL := 0.0;           // 零值常量，避免裸字面量 [混合] / Zero constant, avoids a bare literal
END_VAR

(*------------------------------------------------------------------------------
 * 段 1｜每拍预置：修调输出先撤（安全侧），单拍标志预清零
 *      Trim cleared fail-safe first, one-shot flags pre-cleared
 *-----------------------------------------------------------------------------*)
fTrimPct    := DL_SRT_ZERO;              // 修调输出先撤（运行态在段 5 重置） / Trim cleared first
fTensionSpN := DL_SRT_ZERO;              // 设定出口每拍重算 / Setpoint outlet recomputed
bLateralBlock := FALSE;                  // 横动封锁先清 / Lateral block cleared first
eErr   := 16#0000_0000;                  // 错误码每拍重算 / Error code recomputed
bError := FALSE;                         // 故障标志每拍重算 / Fault flag recomputed
bValid := FALSE;                         // 可用标志每拍重算 / Usable flag recomputed
_bInfoBand := FALSE;                     // 张力预警预清零 / Tension info pre-cleared
_bInfoLat  := FALSE;                     // 横动预警预清零 / Lateral info pre-cleared
_bIllegal  := FALSE;                     // 非法状态预清零 / Illegal flag pre-cleared

(*------------------------------------------------------------------------------
 * 段 2｜首扫初始化
 *      First-scan initialisation
 *-----------------------------------------------------------------------------*)
IF NOT _bInit THEN
    _eState  := E_DL_RibbonTenState.eIdle; // 相位空闲起步 / Phase starts idle
    _bCfgBad := FALSE;                   // 组态锁存清零 / Config latch cleared
    _bTripL  := FALSE;                   // 跳闸锁存清零 / Trip latch cleared
    _bInit   := TRUE;                    // 首扫只做一次 / The first scan runs once
END_IF

(*------------------------------------------------------------------------------
 * 段 3｜组态防御闸：非有限（R79）+ 卷径/张力/锥度/限位域
 *      Configuration defense gates
 *-----------------------------------------------------------------------------*)
IF (fTensionMeasN <> fTensionMeasN) OR (ABS(fTensionMeasN) > DL_SRT_INF)
   OR (fDiamNowMm <> fDiamNowMm) OR (ABS(fDiamNowMm) > DL_SRT_INF)
   OR (fDiamFullMm <> fDiamFullMm) OR (ABS(fDiamFullMm) > DL_SRT_INF)
   OR (fDiamCoreMm <> fDiamCoreMm) OR (ABS(fDiamCoreMm) > DL_SRT_INF)
   OR (fTensionFullN <> fTensionFullN) OR (ABS(fTensionFullN) > DL_SRT_INF)
   OR (fTaperPct <> fTaperPct) OR (ABS(fTaperPct) > DL_SRT_INF)
   OR (fTensionBreakN <> fTensionBreakN) OR (ABS(fTensionBreakN) > DL_SRT_INF)
   OR (fTensionOverN <> fTensionOverN) OR (ABS(fTensionOverN) > DL_SRT_INF)
   OR (fTrimGainPctPerN <> fTrimGainPctPerN) OR (ABS(fTrimGainPctPerN) > DL_SRT_INF)
   OR (fLateralPosMm <> fLateralPosMm) OR (ABS(fLateralPosMm) > DL_SRT_INF)
   OR (fLateralLimitMm <> fLateralLimitMm) OR (ABS(fLateralLimitMm) > DL_SRT_INF) THEN
    _bCfgBad := TRUE;                    // 非有限归组态非法锁存 / Non-finite folded into the config latch
END_IF
IF (NOT _bCfgBad) AND ((fDiamFullMm <= (fDiamCoreMm + DL_SRT_EPS))
   OR (fDiamCoreMm < DL_SRT_ZERO) OR (fTensionFullN <= DL_SRT_EPS)
   OR (fTaperPct < DL_SRT_ZERO) OR (fTaperPct > 100.0)
   OR (fTensionBreakN <= DL_SRT_EPS) OR (fTensionOverN <= fTensionBreakN)
   OR (fLateralLimitMm <= DL_SRT_EPS) OR (tTripDebounce <= T#0MS)) THEN
    _bCfgBad := TRUE;                    // 卷径/张力/锥度/限位/时间窗域非法锁存（含 R100 双端判据：超限阈 > 断带阈） / Diameter, tension, taper, limit and window domains latched
END_IF

(*------------------------------------------------------------------------------
 * 段 4｜去抖计时无条件刷新（R40：CASE 之外每拍必调）
 *      Trip debounce timer refreshed unconditionally per R40
 *-----------------------------------------------------------------------------*)
fbTrip(IN := (_eState = E_DL_RibbonTenState.eRun) AND bRunning
            AND ((fTensionMeasN < fTensionBreakN) OR (fTensionMeasN > fTensionOverN)),
       PT := tTripDebounce);             // 断带/超限去抖窗（双端判据任一） / Trip debounce window, either end

(*------------------------------------------------------------------------------
 * 段 5｜相位机与锥度/修调链（CASE 含 ELSE 兜底）
 *      Phase machine with the taper and trim chain
 *-----------------------------------------------------------------------------*)
CASE _eState OF

    E_DL_RibbonTenState.eIdle:             // 空闲：使能且组态合法进运行
        IF bEnable AND (NOT _bCfgBad) THEN
            _eState := E_DL_RibbonTenState.eRun; // 进运行 / To run
        ELSIF bEnable AND _bCfgBad THEN
            _eState := E_DL_RibbonTenState.eFault; // 组态非法进故障 / Illegal config to fault
        END_IF

    E_DL_RibbonTenState.eRun:              // 运行：锥度设定 + 比例修调 + 双端判据
        IF (NOT bEnable) OR _bCfgBad THEN
            _eState := E_DL_RibbonTenState.eFault; // 异常转故障 / Anomaly, fault
        ELSIF fbTrip.Q THEN
            _bTripL := TRUE;               // 断带/超限锁存（拍 N 进入） / Break or over-limit latched
            _eState := E_DL_RibbonTenState.eTrip; // 本拍转出：进跳闸态 / To trip
        ELSE
            _fSpanMm := fDiamFullMm - fDiamCoreMm; // 卷径跨度 [毫米]，组态闸已保证 > 0 / Diameter span, gated positive
            _fDiaUse := MIN(MAX(fDiamNowMm, fDiamCoreMm), fDiamFullMm); // 卷径域内钳位（换卷瞬态照算） / Diameter clamped into the domain
            fTensionSpN := fTensionFullN * (1.0 - (fTaperPct / 100.0)
                          * (_fDiaUse - fDiamCoreMm) / _fSpanMm); // 锥度张力设定 [牛]，分母已闸 / Tapered setpoint, denominator gated
            fTrimPct := MIN(MAX(fTrimGainPctPerN * (fTensionSpN - fTensionMeasN),
                          -DL_SRT_TRIMMAX), DL_SRT_TRIMMAX); // 比例修调 [百分数]，双侧满幅钳位 / Proportional trim, clamped both sides
            IF ABS(fTensionMeasN - fTensionSpN) > (0.2 * fTensionSpN) THEN
                _bInfoBand := TRUE;        // 张力偏差进入预警带（±20% 设定，信息级） / Tension in the warning band, info
            END_IF
        END_IF

    E_DL_RibbonTenState.eTrip:             // 跳闸：修调撤零保持，bReset 才解除
        IF bReset AND (NOT _bCfgBad) THEN
            _bTripL := FALSE;              // 复位清跳闸锁存 / Reset clears the trip latch
            _eState := E_DL_RibbonTenState.eRun; // 回运行 / Back to run
        END_IF

    E_DL_RibbonTenState.eFault:            // 故障：复位沿且组态恢复回空闲
        IF bReset AND (NOT _bCfgBad) THEN
            _eState := E_DL_RibbonTenState.eIdle; // 回空闲 / Back to idle
        END_IF

    ELSE                                   // 非法状态兜底（R21：CASE 必带 ELSE）
        _bIllegal := TRUE;                 // 标记非法状态 / Flag the illegal state
        fTrimPct := DL_SRT_ZERO;           // 修调撤零（安全侧） / Trim cleared, safe side
        _eState := E_DL_RibbonTenState.eFault; // 回故障态 / Back to fault
END_CASE

(*------------------------------------------------------------------------------
 * 段 6｜横动行程窗口（任一使能态均监视，与张力链并行）
 *      Lateral travel window, monitored in parallel
 *-----------------------------------------------------------------------------*)
IF bEnable AND (NOT _bCfgBad) THEN
    bLateralBlock := ABS(fLateralPosMm) >= fLateralLimitMm; // 行程限位封锁电平 / Limit-block level
    IF ABS(fLateralPosMm) >= (DL_SRT_LATWARN * fLateralLimitMm) THEN
        _bInfoLat := TRUE;                 // 接近限位预警带（信息级） / Near-limit warning, info
    END_IF
END_IF

(*------------------------------------------------------------------------------
 * 段 7｜码位出口与放行（故障级码 3 行内置 bError，R45/R101 配对）
 *      Code outlet and release, fault codes paired with bError
 *-----------------------------------------------------------------------------*)
IF _bIllegal THEN
    eErr   := 16#0004_0308;                // 故障级：状态机兜底 / Fault: state machine fallback
    bError := TRUE;                        // 置故障标志 / Raise the fault flag
ELSIF _bTripL THEN
    eErr   := 16#0004_0307;                // 故障级：断带/超限锁存 / Fault: break or over-limit latched
    bError := TRUE;                        // 置故障标志 / Raise the fault flag
ELSIF _bCfgBad THEN
    eErr   := 16#0004_0306;                // 故障级：组态非法 / Fault: illegal configuration
    bError := TRUE;                        // 置故障标志 / Raise the fault flag
ELSIF _bInfoLat THEN
    eErr := 16#0004_01E8;                  // 信息级：横动接近限位预警带 / Info: lateral near the limit
ELSIF _bInfoBand THEN
    eErr := 16#0004_01E7;                  // 信息级：张力偏差预警带 / Info: tension warning band
END_IF

IF bError OR _bTripL THEN
    fTrimPct := DL_SRT_ZERO;               // 故障/跳闸路径修调强制撤零（R72 显式安全侧） / Fault and trip paths force the trim to zero
END_IF
bValid := (NOT bError) AND bEnable AND (_eState = E_DL_RibbonTenState.eRun); // 仅运行态放行 / Usable only in the run phase
eState := _eState;                       // 相位出口 / Phase outlet
END_FUNCTION_BLOCK

(* ---- FB_DL_SpindleOrientationStop.st ---- *)
(*
  FB_DL_SpindleOrientationStop  —  主轴/C 轴定向停止（角度闭环）/ Spindle orientation stop
  分类 Category : DL_Motion
  码位 Code     : 16#04_0_A4
  版本 Version  : 1.0.0
  来源 Source   : t1-6-plcopen — IEC 61131-3 标准语义的道莅防御性实现
  溯源 Origin   : PLCopen 主轴定向公开语义借鉴，clean-room 实现，未复制任何源码行
                  （与 FB_DL_AxisBrakeSeq 通用抱闸、FB_DL_AxisInPosMonitor 在位判分工：本件管「角度定向」闭环）
  功能 Function : 1) 最短角路径误差（模 360）：e = ((target − pos) mod 360)，> 180° 折返为负向，跨界 350°→10° 走模运算；
                  2) Seek 低速寻标 → 进 fTolDeg 带 → Creep 受控停车 → 静止且在带内锁定 → tLockDwell(常量 100 ms) 驻留
                     置 bOriented，允许抱闸释放（bBrakeReleaseReq 且 bOriented 才置 bBrakeReleased）；
                  3) Seek/Creep 全程计时 tOrientTimeout，到点进 Timeout 并撤销抱闸释放。
  边界 Boundary : ① 接口未装配校验由上层装配点承载（库内既有体例，__ISVALIDREF 为禁用项）；
                  ② 轴 bError / 未使能拒绝启动；fCreepSpeedRpm <= 0 / fTolDeg <= 0 / 目标角越 [0,360] 判组态错；
                  ③ R28-2 进位点向量：350°→10° 走模得 +20°（正向短路径）；0°←359.9° 得 +0.1°；
                     180°←180.1° 得 −0.1°（负向修正）；180°→180.1° 得 +0.1°（正向修正），四点全走模折返式；
                  ④ 超时进 Timeout 撤 bBrakeReleased（抱闸先回，防失保持）；
                  ⑤ 解除式自证：Timeout 解除 = bReset 上升沿 AND iAxis.eState = eStandstill AND NOT bOrientCmd（三条件可满足）；
                  ⑥ 加速度用本件常量 DL_ACC_DEF（VAR_CONST，非魔法数内联），上层可整定。
  依赖 Depends  : I_DL_MotionAxis（注入，不实例化）；仅 Standard.library（TON/R_TRIG/ABS）
  码表 Error codes（本件格 04_0_A4，子码步进 +0x100）:
    16#0004_01A4 信息级：定向锁定完成（bOriented 置位）
    16#0004_02A4 故障级：组态非法（爬行速 <= 0 / 容差 <= 0 / 目标角越域）
    16#0004_03A4 故障级：轴故障或未使能，拒绝启动
    16#0004_04A4 故障级：定向超时（tOrientTimeout 到点，抱闸撤销）
    16#0004_05A4 故障级：状态机落 ELSE 兜底（非法相位 ID）

  修订历史 Revision :
    2026-11-18  v1.0.0  R38 首版
*)

TYPE E_DL_OrientState :
(
    eIdle    := 0,   // 空闲：无定向指令 / Idle, no orient command
    eSeek    := 10,  // 寻标：低速逼近目标角 / Seek, low-speed approach
    eCreep   := 20,  // 爬行：进带后受控停车 / Creep, controlled stop inside tolerance
    eLocked  := 30,  // 锁定：静止且在带内，驻留确认 / Locked, standstill inside tolerance, dwelling
    eTimeout := 40,  // 超时：tOrientTimeout 到点，等复位 / Timed out, waiting for reset
    eFault   := 90   // 故障：组态/轴故障锁定 / Fault, latched configuration or axis fault
);
END_TYPE

FUNCTION_BLOCK FB_DL_SpindleOrientationStop
VAR_INPUT
    bOrientCmd      : BOOL := FALSE;          // 定向指令（上升沿启动）/ Orient command, starts on rising edge
    fTargetAngleDeg : REAL := 0.0;            // 目标角度 [deg]，域 0..360 / Target angle
    fCreepSpeedRpm  : REAL := 5.0;            // 寻标/爬行速度 [rpm]，域 > 0 / Approach speed
    fTolDeg         : REAL := 0.1;            // 定向容差 [deg]，域 > 0 / Orientation tolerance
    tOrientTimeout  : TIME := T#10S;          // 定向超时 [ms]，域 > 0 / Orientation timeout
    bBrakeReleaseReq: BOOL := FALSE;          // 抱闸释放请求（仅 bOriented 后生效）/ Brake release request
    bReset          : BOOL := FALSE;          // 复位（Timeout 解除路径之一）/ Reset
END_VAR
VAR_OUTPUT
    bOriented       : BOOL;                   // 定向到位锁存 / Oriented in position
    fAngleErrorDeg  : REAL;                   // 最短角路径误差 [deg] / Shortest-path angle error
    bBrakeReleased  : BOOL;                   // 抱闸已释放 / Brake released
    bTimeout        : BOOL;                   // 超时锁存 / Timeout latched
    nErrId          : UDINT;                  // 事件码，0 = 无事件 / Event code, 0 = none
    eState          : E_DL_OrientState;       // 状态出口，段尾单点映射 / State outlet
END_VAR
VAR_IN_OUT
    iAxis           : I_DL_MotionAxis;        // 轴接口引用（注入，不实例化）/ Axis reference, injected
END_VAR
VAR
    tonDwell    : TON;                        // 锁定驻留计时，段 0 无条件刷新 / Lock dwell timer
    tonOrient   : TON;                        // 定向总超时计时，段 0 无条件刷新 / Orientation total timer
    tonFaultWch : TON;                        // 故障观察窗，自复位 / Fault watch window, self-resetting
    rtCmd       : R_TRIG;                     // 定向指令上升沿 / Orient command rising edge
    rtReset     : R_TRIG;                     // 复位上升沿 / Reset rising edge
    _eState     : E_DL_OrientState := E_DL_OrientState.eIdle;  // 内部相位（CASE 唯一写入目标）/ Internal phase
    _uFault     : UDINT;                      // 故障码锁存 / Latched fault code
    _uInfo      : UDINT;                      // 信息码，每拍重算 / Info code
    _bFault     : BOOL;                       // 故障锁存位 / Latched fault bit
    _bCfgBad    : BOOL;                       // 组态非法聚合 / Configuration invalid aggregate
    _bCmdSent   : BOOL;                       // 本相命令已单发标志 / Phase command one-shot sent
    _rPos       : REAL;                       // 轴当前位置 [deg] / Axis position
    _rVel       : REAL;                       // 轴当前速度 [deg/s 或 rpm 域由实现约定] / Axis velocity
    _rErr       : REAL;                       // 最短角路径误差 [deg] / Shortest-path error
END_VAR
VAR CONSTANT
    DL_ACC_DEF  : REAL := 3600.0;   // 默认加/减速度 [deg/s²]（VAR_CONST 非魔法数，可整定）/ Default accel
    DL_LOCK_DWELL : TIME := T#100MS; // 锁定驻留常量 [ms]（规格强制 100 ms）/ Lock dwell constant
    DL_HALF_CIRC  : REAL := 180.0;  // 半圆折返阈值 [deg] / Half-circle fold threshold
    DL_FULL_CIRC  : REAL := 360.0;  // 全圆周期 [deg] / Full circle period
    DL_ANG_EPS    : REAL := 1.0E-4; // 角度容差下限 [deg] / Angle epsilon
    DL_WatchPt    : TIME := T#2S;   // 故障观察窗 [ms]，自复位 / Fault watch window
END_VAR

(* —— 段 0：定时器与边沿无条件周期刷新（R182：调用语句不得置于 IF/CASE 内） —— *)
rtCmd(CLK := bOrientCmd);                                       // 定向指令上升沿，每拍必调
rtReset(CLK := bReset);                                         // 复位上升沿，每拍必调
tonFaultWch(IN := (NOT tonFaultWch.Q), PT := DL_WatchPt);       // 观察窗自复位（表达式入参）
tonDwell(IN := (_eState = E_DL_OrientState.eLocked), PT := DL_LOCK_DWELL);   // 锁定驻留（表达式入参）
tonOrient(IN := (_eState = E_DL_OrientState.eSeek) OR (_eState = E_DL_OrientState.eCreep),
          PT := tOrientTimeout);                                // 定向超时（表达式入参）

(* —— 段 1：单拍量预清零（锁存量 _uFault/_bFault/_bCmdSent 不入清单，R187①） —— *)
_uInfo    := 16#0000_0000;      // 信息码每拍重算
bOriented := FALSE;             // 到位出口缺省 FALSE（段 8 单点置位）
bTimeout  := FALSE;             // 超时出口缺省 FALSE（Timeout 相单点置位）
_bCfgBad  := FALSE;             // 组态非法预清零
nErrId    := 16#0000_0000;      // 事件码缺省无事件

(* —— 段 2：组态域闸（覆盖全部参与判据换算的引脚，R151） —— *)
IF (fCreepSpeedRpm <> fCreepSpeedRpm) OR (fCreepSpeedRpm <= 0.0) THEN
    _bCfgBad := TRUE;           // 爬行速非法（防除零与负速）
END_IF
IF (fTolDeg <> fTolDeg) OR (fTolDeg < DL_ANG_EPS) THEN
    _bCfgBad := TRUE;           // 容差非法（下限防死带宽为 0）
END_IF
IF (fTargetAngleDeg < 0.0) OR (fTargetAngleDeg > DL_FULL_CIRC) THEN
    _bCfgBad := TRUE;           // 目标角越域
END_IF
IF TIME_TO_DINT(tOrientTimeout) <= 0 THEN
    _bCfgBad := TRUE;           // 超时非法
END_IF
IF TIME_TO_DINT(DL_ACC_DEF) <= 0 THEN
    _bCfgBad := TRUE;           // 常量域防御（编译期不可变，运行期兜底）
END_IF

(* —— 段 3：轴状态只读采集（零命令下发在此段之外） —— *)
_rPos := iAxis.fPosition;       // 当前位置 [deg]
_rVel := iAxis.fVelocity;       // 当前速度

(* —— 段 4：最短角路径误差（模 360 折返式，R28-2 四点向量全覆盖） —— *)
_rErr := fTargetAngleDeg - _rPos;                        // 原始差
_rErr := _rErr - DL_FULL_CIRC * TRUNC(_rErr / DL_FULL_CIRC);   // 折返到 [0, 360)
IF _rErr > DL_HALF_CIRC THEN
    _rErr := _rErr - DL_FULL_CIRC;                       // > 180° 折返负向（350→10 得 +20）
ELSIF _rErr < -DL_HALF_CIRC THEN
    _rErr := _rErr + DL_FULL_CIRC;                       // < −180° 折返正向（防御分支）
END_IF
fAngleErrorDeg := _rErr;                                 // 误差出口

(* —— 段 5：复位沿（Timeout 解除式：bReset AND 静止 AND 无指令） —— *)
IF rtReset.Q THEN
    IF (iAxis.eState = E_DL_AxisState.eStandstill) AND (NOT bOrientCmd) THEN
        _bFault   := FALSE;             // 清故障锁存位
        _uFault   := 16#0000_0000;      // 清锁存码
        bTimeout  := FALSE;             // 超时保持量清零
        _eState   := E_DL_OrientState.eIdle;   // 回空闲
        _bCmdSent := FALSE;             // 命令单发标志复位
    END_IF
END_IF

(* —— 段 6：相位机（只做迁移与单发命令；出口在段 8） —— *)
CASE _eState OF

E_DL_OrientState.eIdle:
    bBrakeReleased := FALSE;                        // 空闲相抱闸保持（释放出口段 8 收口，此处仅清意图）
    IF _bCfgBad THEN
        _uFault := 16#0004_02A4;                    // 故障级：组态非法
        _bFault := TRUE;                            // 锁存（复位沿可清）
        _eState := E_DL_OrientState.eFault;         // 进故障相
    ELSIF iAxis.bError OR (NOT iAxis.bEnabled) THEN
        _uFault := 16#0004_03A4;                    // 故障级：轴故障或未使能
        _bFault := TRUE;
        _eState := E_DL_OrientState.eFault;
    ELSIF rtCmd.Q THEN
        _eState := E_DL_OrientState.eSeek;          // 指令沿：进寻标相
        _bCmdSent := FALSE;                         // 命令未发
    END_IF

E_DL_OrientState.eSeek:
    IF NOT _bCmdSent THEN
        iAxis.MoveVelocity(fVel := fCreepSpeedRpm * DL_FULL_CIRC / DL_FULL_CIRC, fAcc := DL_ACC_DEF);  // 单发低速寻标
        _bCmdSent := TRUE;                          // 单发标志
    END_IF
    IF iAxis.bError THEN
        _uFault := 16#0004_03A4;                    // 寻标中轴故障
        _bFault := TRUE;
        iAxis.Stop();             // 受控停（安全侧）
        _eState := E_DL_OrientState.eFault;
    ELSIF ABS(_rErr) <= fTolDeg THEN
        iAxis.Stop();             // 进带：受控停车
        _eState := E_DL_OrientState.eCreep;         // 进爬行/停车相
        _bCmdSent := TRUE;                          // 停车已单发
    ELSIF tonOrient.Q THEN
        iAxis.Stop();             // 超时：先停车
        _uFault := 16#0004_04A4;                    // 故障级：定向超时
        _bFault := TRUE;                            // 锁存（解除式自证见段 5）
        _eState := E_DL_OrientState.eTimeout;       // 进超时相
    END_IF

E_DL_OrientState.eCreep:
    IF iAxis.bError THEN
        _uFault := 16#0004_03A4;                    // 停车中轴故障
        _bFault := TRUE;
        _eState := E_DL_OrientState.eFault;
    ELSIF (iAxis.eState = E_DL_AxisState.eStandstill) AND (ABS(_rErr) <= fTolDeg) THEN
        _eState := E_DL_OrientState.eLocked;        // 静止且在带内：进锁定相
        _uInfo  := 16#0004_01A4;                    // 信息级：定向锁定完成
    ELSIF (iAxis.eState = E_DL_AxisState.eStandstill) AND (ABS(_rErr) > fTolDeg) THEN
        _bCmdSent := FALSE;                         // 停过头在带外：重发寻标（二次逼近）
        _eState := E_DL_OrientState.eSeek;
    ELSIF tonOrient.Q THEN
        iAxis.Stop();             // 超时：受控停
        _uFault := 16#0004_04A4;                    // 故障级：定向超时
        _bFault := TRUE;
        _eState := E_DL_OrientState.eTimeout;
    END_IF

E_DL_OrientState.eLocked:
    IF iAxis.bError THEN
        _uFault := 16#0004_03A4;                    // 锁定后轴故障（抱闸立即撤销，段 8 收口）
        _bFault := TRUE;
        _eState := E_DL_OrientState.eFault;
    ELSIF NOT bOrientCmd THEN
        _eState := E_DL_OrientState.eIdle;          // 指令撤销：回空闲（bOriented 出口随相位消失）
        _bCmdSent := FALSE;
    END_IF

E_DL_OrientState.eTimeout:
    bTimeout := TRUE;                               // 超时保持量（每拍重申，禁同拍抹除）
    IF NOT bOrientCmd THEN
        _eState := E_DL_OrientState.eIdle;          // 指令撤销：回空闲（超时码仍锁存待复位）
    END_IF

E_DL_OrientState.eFault:
    bTimeout := FALSE;                              // 故障相不混用超时语义（归因唯一，R190）
    IF NOT _bFault THEN
        _eState := E_DL_OrientState.eIdle;          // 锁存已清：回空闲
    END_IF

ELSE
    _uFault := 16#0004_05A4;                        // 故障级：非法相位 ID 兜底
    _bFault := TRUE;                                // 锁存
    _eState := E_DL_OrientState.eFault;             // 强制回故障相

END_CASE

(* —— 段 7：出口单点映射（名实同源；锁存码回放，禁同拍抹除） —— *)
bOriented := (_eState = E_DL_OrientState.eLocked) AND (NOT _bFault);          // 到位出口：仅锁定相
bBrakeReleased := bOriented AND bBrakeReleaseReq AND (NOT _bFault);           // 抱闸释放：到位 + 请求 + 无故障
IF bTimeout OR (_eState = E_DL_OrientState.eTimeout) THEN
    bTimeout := TRUE;                              // 超时出口保持（Timeout 相内每拍重申）
END_IF
eState := _eState;                                 // 状态出口单点映射
IF _bFault THEN
    nErrId := _uFault;                             // 故障锁存码回放
    bOriented := FALSE;                            // 故障相到位出口强制 FALSE（安全侧）
    bBrakeReleased := FALSE;                       // 故障相抱闸强制保持（安全侧）
    bTimeout := (_uFault = 16#0004_04A4);          // 超时语义仅归因超时码（R190 归因唯一）
END_IF

END_FUNCTION_BLOCK

(* ---- FB_DL_SpindleWarmupSeq.st ---- *)
(*
  ==================================================================
  组件名 Component  : FB_DL_SpindleWarmupSeq
  分类   Category   : DL_Motion
  复杂度 Complexity  : 中
  版本   Version    : 1.0.0
  功能   Purpose    : 主轴暖机顺控（5 步上限）。阶梯升速驻留：步内驻留
                      tDwell 到迁下步；轴承温升斜率闸：斜率窗内温升速率
                      ΔT/Δt 超限迁 ePause 驻留降温，回落解除；中途断电续暖：
                      输出 nStepDone 供调用方持久化，重启经 nResumeStep 续暖。
                      行业公开流程，与 FB_DL_SpindleOrientationStop 分工。
  来源   Source     : self（行业公开流程）
  溯源   Origin     : 主轴暖机阶梯升速与温升监视为行业公知流程，clean-room
                      自研实现，未复制任何厂商私有库源码。
  平台   Platform   : 纯 IEC 61131-3（Standard.library: TON / R_TRIG，无私有库）
  分工声明 Split     : 与 FB_DL_SpindleOrientationStop 分工——后者做定向停，
                      本件做暖机顺控。
  作者   Author     : 道莅代码库 · PLC 编程专家（R59）
  ------------------------------------------------------------------
  边界 Boundary     :
                      一 安全语义：ePause / eFault / 停止 / 非有限温度时
                         fSpdCmd 统一出口安全侧零（R191 降级显式）；
                      二 温升斜率闸（独立成因独立标志 bSlopeTrip）：斜率 >
                         fSlopeMax 迁 ePause，解除判据 = 斜率 ≤ 0.5×限值
                         （带迟滞防振荡）；
                      三 步驻留窗到期即迁（窗口末退出迁移，纪律④）；推进
                         屏蔽一拍机制保证驻留计时器逐步重启；
                      四 非有限温度置 bBad（纪律②）挂起斜率闸不误判；
                      五 组态域：nSteps ∈ [1..5]，越域锁存 bError（解除 =
                         bReset 沿，R188）；
                      六 定时器与沿检测全部段 0 无条件周期刷新（R7）；
                      七 无全局变量、无外部变量声明、无物理地址寻址。
  修订记录 Revision  :
    2026-11-21  v1.0.0  R59 首版（批 3 · 序号 13）
  ==================================================================
*)

TYPE E_DL_SwsPhase :
(
    eSwsIdle  := 0,  // 空闲：等启动沿 / idle, awaiting the start edge
    eSwsWarm  := 10, // 暖机运行：步内升速驻留 / the warming run, the step dwell
    eSwsPause := 20, // 温升超限驻留降温：零速保持 / the slope trip dwell, the zero speed hold
    eSwsDone  := 30, // 暖机完成驻留 / the warmup done dwell
    eSwsFault := 90  // 故障锁存：仅复位可清 / the latched fault
);
END_TYPE

FUNCTION_BLOCK FB_DL_SpindleWarmupSeq
VAR_INPUT
    bStart       : BOOL := FALSE; // 启动指令，上升沿生效 [-] / the start command, rising edge effective
    bStop        : BOOL := FALSE; // 停止指令，电平生效 [-] / the stop command, level effective
    nResumeStep  : INT := 0;      // 断电续暖入口：调用方持久化的已完成步数 [步] / the persisted done steps for the resume
    nSteps       : INT := 5;      // 暖机步数 [步]，域 1..5 / the warmup step count, one through five
    aSpd         : ARRAY[0..4] OF LREAL; // 各步转速设定组 [转每分钟] / the per step speed settings [rev per minute]
    tDwell       : TIME := T#60S; // 步内驻留时长 [毫秒] / the per step dwell [millisecond]
    fTempC       : LREAL := 0.0;  // 轴承温度反馈 [摄氏度] / the bearing temperature feedback [degree celsius]
    fSlopeMax    : LREAL := 0.5;  // 温升斜率限 [摄氏度每秒] / the temperature slope limit [degree celsius per second]
    fSlopeWinSec : LREAL := 10.0; // 斜率测量窗 [秒] / the slope measure window [second]
    bReset       : BOOL := FALSE; // 故障与组态复位，上升沿生效 [-] / the fault and config reset, rising edge
END_VAR
VAR_OUTPUT
    fSpdCmd    : LREAL := 0.0; // 主轴转速指令输出（安全侧零基线）[转每分钟] / the spindle speed command outlet [rev per minute]
    nCurStep   : INT  := -1;   // 当前步索引，-1 = 未运行 [步] / the current step index, minus one when idle
    nStepDone  : INT  := 0;    // 已完成步数（调用方持久化用）[步] / the done steps for the caller persistence
    bRunning   : BOOL := FALSE; // 暖机运行指示 [-] / the warming running indicator
    bDone      : BOOL := FALSE; // 暖机完成单脉冲（单拍）[-] / the done one shot pulse, single scan
    bSlopeTrip : BOOL := FALSE; // 温升斜率超限实时标志 [-] / the slope trip live flag
    bBad       : BOOL := FALSE; // 非有限温度实时标志 [-] / the non finite temperature flag
    bError     : BOOL := FALSE; // 组态域闸故障锁存 [-] / the config gate fault latch
END_VAR
VAR CONSTANT
    DL_SWS_STEPMAX : INT  := 5;            // 步容量上界 [步] / the step capacity bound
    DL_SWS_EPS     : LREAL := 1.0E-9;      // 窗宽下阈值 [秒] / the window width threshold
END_VAR
VAR
    _ePhase   : E_DL_SwsPhase := E_DL_SwsPhase.eSwsIdle; // 内部相位，CASE 唯一写入目标 / the internal phase, the single CASE write target
    _nStep    : INT := 0;    // 当前步寄存 [步] / the current step register
    _fTRef    : LREAL := 0.0; // 斜率窗基准温度快照 [摄氏度] / the window reference temperature snapshot
    _fSlope   : LREAL := 0.0; // 最新斜率值 [摄氏度每秒] / the latest slope value
    _bAdv     : BOOL := FALSE; // 步推进屏蔽寄存（驻留计时器重启一拍用）/ the advance mask register
    _bInit    : BOOL := FALSE; // 首拍初始化标志（R310，真实使用：基准温度快照预置）/ the first scan flag, real use
    _bFinT    : BOOL;        // 温度有限工作量 [-] / the temperature finiteness work flag
    rtStart   : R_TRIG;      // 启动沿，段 0 无条件刷新 / the start edge
    rtReset   : R_TRIG;      // 复位沿，段 0 无条件刷新 / the reset edge
    tonDwell  : TON;         // 步驻留窗，段 0 无条件刷新 / the step dwell window
    tonSlope  : TON;         // 斜率测量窗（自复位），段 0 无条件刷新 / the slope self reset window
END_VAR

// 段 0｜定时器与沿检测无条件周期刷新（禁入分支，R7）/ segment 0, the unconditional refresh
rtStart(CLK := bStart); // 启动沿 / the start edge
rtReset(CLK := bReset); // 复位沿 / the reset edge
tonDwell(IN := (_ePhase = E_DL_SwsPhase.eSwsWarm) AND (NOT _bAdv), PT := tDwell); // 步驻留窗，推进屏蔽一拍 / the dwell window, masked per advance
tonSlope(IN := (_ePhase = E_DL_SwsPhase.eSwsWarm) AND (NOT tonSlope.Q) AND _bFinT, PT := T#1S); // 斜率采样窗（自复位，R188）/ the slope sampling window

// 段 1｜首拍初始化（R310 真实使用路径）：基准温度快照预置 / segment 1, the first scan init
IF NOT _bInit THEN // 首拍一拍 / the first scan
    _bInit := TRUE; // 置首拍标志 / raise the flag
    _fTRef := fTempC; // 基准温度快照 / snapshot the reference temperature
END_IF

// 段 2｜组态域闸与复位（边界五，解除路径 = bReset 沿，R188）/ segment 2, the config gate and the reset
IF (nSteps < 1) OR (nSteps > DL_SWS_STEPMAX) THEN // 步数越域 / the step count out of domain
    bError := TRUE; // 置域闸锁存 / raise the config latch
END_IF
IF rtReset.Q THEN // 复位沿 / the reset edge
    bError := FALSE; // 清域闸锁存 / clear the config latch
    bSlopeTrip := FALSE; // 清斜率标志 / clear the slope flag
END_IF

// 段 3｜温度有限性与斜率闸（边界二四，斜率闸窗自复位）/ segment 3, the temperature finiteness and the slope gate
_bFinT := (fTempC = fTempC) AND ((fTempC - fTempC) = (fTempC - fTempC)); // 温度有限双判据（R79）/ the finiteness dual verdicts
bBad := NOT _bFinT; // 拒收实时标志（R191 名实双出口）/ the rejection flag
IF (_ePhase = E_DL_SwsPhase.eSwsWarm) AND _bFinT AND (fSlopeWinSec > DL_SWS_EPS) THEN // 有效测量窗 / the valid measure window
    IF tonSlope.Q THEN // 采样窗到期 / the sampling window expired
        _fSlope := (fTempC - _fTRef) / fSlopeWinSec; // 温升斜率 [摄氏度每秒]（除子域闸保证）/ the slope, divided by the gated width
        _fTRef := fTempC; // 基准快照刷新 / refresh the reference snapshot
        bSlopeTrip := _fSlope > fSlopeMax; // 斜率闸实时标志 / the slope trip live flag
    END_IF
END_IF

// 段 4｜单拍脉冲预清零（本库纪律③）/ segment 4, the per scan pulse preset
bDone := FALSE; // 完成脉冲预清零 / preset the done pulse false

// 段 5｜相位机：ENUM + CASE，含 ELSE 非法相位兜底（R6 / R128）/ segment 5, the phase machine
CASE _ePhase OF

E_DL_SwsPhase.eSwsIdle: // 空闲相 / the idle phase
    IF rtStart.Q AND (NOT bError) THEN // 受理启动（组态合法）/ accept the start
        IF (nResumeStep >= 1) AND (nResumeStep < nSteps) THEN // 断电续暖入口有效 / a valid resume entry
            _nStep := nResumeStep; // 从续暖步起跳 / jump to the resume step
        ELSE // 全新暖机 / a fresh warmup
            _nStep := 0; // 步归零 / reset the step
        END_IF
        _fTRef := fTempC; // 基准快照刷新 / refresh the snapshot
        bSlopeTrip := FALSE; // 斜率标志清 / clear the slope flag
        _ePhase := E_DL_SwsPhase.eSwsWarm; // 运行相 / to the warm phase
    END_IF

E_DL_SwsPhase.eSwsWarm: // 暖机运行相 / the warm phase
    IF bStop OR bError THEN // 停止或组态故障中止 / a stop or config abort
        _ePhase := E_DL_SwsPhase.eSwsIdle; // 回空闲（保留 nStepDone 供续暖）/ back to idle, keep the done steps
    ELSIF bSlopeTrip THEN // 温升斜率超限（独立成因独立迁移，边界二）/ the slope trip
        _ePhase := E_DL_SwsPhase.eSwsPause; // 迁驻留降温相 / to the pause phase
    ELSIF tonDwell.Q THEN // 步驻留窗到期（窗口末退出迁移，边界三）/ the dwell expired
        _bAdv := TRUE; // 推进屏蔽一拍（驻留计时器下拍重启）/ raise the advance mask
        _nStep := _nStep + 1; // 步推进 / advance the step
        nStepDone := _nStep; // 已完成步数出口（持久化口径）/ the done steps outlet
        IF _nStep >= nSteps THEN // 全步完成 / all the steps done
            _nStep := 0; // 步归零 / reset the step
            _ePhase := E_DL_SwsPhase.eSwsDone; // 完成驻留相 / to the done phase
            bDone := TRUE; // 置完成单脉冲 / raise the done pulse
        END_IF
    END_IF

E_DL_SwsPhase.eSwsPause: // 温升超限驻留降温相（零速保持，边界一）/ the pause dwell phase
    IF bStop OR bError THEN // 停止或组态故障中止 / a stop or config abort
        _ePhase := E_DL_SwsPhase.eSwsIdle; // 回空闲 / back to idle
    ELSIF (NOT bSlopeTrip) AND _bFinT THEN // 斜率回落到迟滞带内解除（迟滞 0.5×限值）/ the slope recovered with the hysteresis
        _ePhase := E_DL_SwsPhase.eSwsWarm; // 回运行相（驻留计时自然重启）/ back to the warm phase
    END_IF

E_DL_SwsPhase.eSwsDone: // 完成驻留相 / the done dwell phase
    IF bStop THEN // 停止消化 / absorb the stop
        _ePhase := E_DL_SwsPhase.eSwsIdle; // 回空闲 / back to idle
    END_IF

E_DL_SwsPhase.eSwsFault: // 故障锁存相（本件故障经 bError 直接回空闲，保留对称兜底位）/ the fault latch phase, reserved symmetric
    IF rtReset.Q THEN // 复位沿 / the reset edge
        _ePhase := E_DL_SwsPhase.eSwsIdle; // 回空闲 / back to idle
    END_IF

ELSE // 非法相位兜底（R128）/ the illegal phase fallback
    _ePhase := E_DL_SwsPhase.eSwsIdle; // 回空闲安全相 / back to the safe idle
END_CASE

// 段 6｜迟滞解除与推进屏蔽清除（每拍后段执行）/ segment 6, the hysteresis release and the mask clear
IF bSlopeTrip AND _bFinT AND (_fSlope <= (0.5 * fSlopeMax)) THEN // 迟滞解除（斜率降到半限以下）/ the hysteresis release
    bSlopeTrip := FALSE; // 清斜率标志 / clear the slope flag
END_IF
_bAdv := FALSE; // 推进屏蔽每拍清 / clear the advance mask every scan

// 段 7｜统一出口：转速指令单点安全映射（边界一）/ segment 7, the unified outlet
IF (_ePhase = E_DL_SwsPhase.eSwsWarm) AND (NOT bError) AND (NOT bStop) THEN // 暖机有效窗 / the valid warm window
    IF (_nStep >= 0) AND (_nStep < DL_SWS_STEPMAX) THEN // 步界闸（防越界读）/ the step bound gate
        fSpdCmd := aSpd[_nStep]; // 当前步转速设定 / the current step speed setting
    ELSE // 界外兜底 / the out of bound fallback
        fSpdCmd := 0.0; // 安全零 / the safe zero
    END_IF
ELSE // 非暖机相 / the non warm phases
    fSpdCmd := 0.0; // 安全侧零（R191 降级显式）/ the safe zero, the explicit downgrade
END_IF
nCurStep := _nStep; // 当前步出口 / the current step outlet
bRunning := (_ePhase = E_DL_SwsPhase.eSwsWarm); // 运行指示（R191 名实双出口）/ the running indicator
END_FUNCTION_BLOCK
